  movel([0.337067, -0.804925, -2.801835, -1.105629, 1.570796, 1.907863],accel_mss,speed_ms,0,blend_radius_m)
  movel([0.336030, -0.804781, -2.801859, -1.105749, 1.570796, 1.906826],accel_mss,speed_ms,0,blend_radius_m)
  movel([0.330509, -0.802988, -2.802160, -1.107241, 1.570796, 1.901306],accel_mss,speed_ms,0,blend_radius_m)
  movel([0.325271, -0.800769, -2.802530, -1.109089, 1.570796, 1.896067],accel_mss,speed_ms,0,blend_radius_m)
  movel([0.320318, -0.798128, -2.802968, -1.111294, 1.570796, 1.891115],accel_mss,speed_ms,0,blend_radius_m)
  movel([0.315671, -0.795055, -2.803472, -1.113862, 1.570796, 1.886468],accel_mss,speed_ms,0,blend_radius_m)
  movel([0.314088, -0.793737, -2.803687, -1.114965, 1.570796, 1.884885],accel_mss,speed_ms,0,blend_radius_m)
  movel([0.312919, -0.791939, -2.803978, -1.116471, 1.570796, 1.883716],accel_mss,speed_ms,0,blend_radius_m)
  movel([0.312565, -0.790531, -2.804206, -1.117652, 1.570796, 1.883362],accel_mss,speed_ms,0,blend_radius_m)
  movel([0.312427, -0.788928, -2.804463, -1.118997, 1.570796, 1.883224],accel_mss,speed_ms,0,blend_radius_m)
  movel([0.312533, -0.785387, -2.805028, -1.121975, 1.570796, 1.883329],accel_mss,speed_ms,0,blend_radius_m)
  movel([0.314201, -0.771715, -2.807148, -1.133527, 1.570796, 1.884998],accel_mss,speed_ms,0,blend_radius_m)
  movel([0.314322, -0.768078, -2.807696, -1.136615, 1.570796, 1.885118],accel_mss,speed_ms,0,blend_radius_m)
  movel([0.313995, -0.765120, -2.808138, -1.139131, 1.570796, 1.884791],accel_mss,speed_ms,0,blend_radius_m)
  movel([0.313608, -0.764022, -2.808300, -1.140066, 1.570796, 1.884404],accel_mss,speed_ms,0,blend_radius_m)
  movel([0.313044, -0.763237, -2.808416, -1.140736, 1.570796, 1.883841],accel_mss,speed_ms,0,blend_radius_m)
  movel([0.312284, -0.762822, -2.808478, -1.141089, 1.570796, 1.883080],accel_mss,speed_ms,0,blend_radius_m)
  movel([0.311307, -0.762817, -2.808478, -1.141093, 1.570796, 1.882104],accel_mss,speed_ms,0,blend_radius_m)
  movel([0.309324, -0.763465, -2.808383, -1.140541, 1.570796, 1.880120],accel_mss,speed_ms,0,blend_radius_m)
  movel([0.308425, -0.763643, -2.808356, -1.140389, 1.570796, 1.879221],accel_mss,speed_ms,0,blend_radius_m)
  movel([0.307786, -0.763410, -2.808391, -1.140588, 1.570796, 1.878582],accel_mss,speed_ms,0,blend_radius_m)
  movel([0.307584, -0.762203, -2.808569, -1.141618, 1.570796, 1.878380],accel_mss,speed_ms,0,blend_radius_m)
  movel([0.307977, -0.760492, -2.808820, -1.143078, 1.570796, 1.878773],accel_mss,speed_ms,0,blend_radius_m)
  movel([0.309463, -0.754879, -2.809633, -1.147877, 1.570796, 1.880260],accel_mss,speed_ms,0,blend_radius_m)
  movel([0.310630, -0.749455, -2.810405, -1.152529, 1.570796, 1.881426],accel_mss,speed_ms,0,blend_radius_m)
  movel([0.312165, -0.739066, -2.811845, -1.161479, 1.570796, 1.882961],accel_mss,speed_ms,0,blend_radius_m)
  movel([0.312944, -0.729061, -2.813184, -1.170144, 1.570796, 1.883740],accel_mss,speed_ms,0,blend_radius_m)
  movel([0.313326, -0.719178, -2.814462, -1.178749, 1.570796, 1.884122],accel_mss,speed_ms,0,blend_radius_m)
  speed_ms = 0.005
  movel([0.313326, -0.711620, -2.807866, -1.192903, 1.570796, 1.884122],accel_mss,speed_ms,0,blend_radius_m)
  speed_ms = 0.040
  movel([0.305588, -0.730189, -2.805441, -1.176759, 1.570796, 1.876385],accel_mss,speed_ms,0,blend_radius_m)
  speed_ms = 0.005
  movel([0.305588, -0.737993, -2.811991, -1.162406, 1.570796, 1.876385],accel_mss,speed_ms,0,blend_radius_m)
  speed_ms = 0.025
  movel([0.301170, -0.750294, -2.810287, -1.151809, 1.570796, 1.871966],accel_mss,speed_ms,0,blend_radius_m)
  movel([0.298692, -0.756493, -2.809401, -1.146496, 1.570796, 1.869489],accel_mss,speed_ms,0,blend_radius_m)
  movel([0.296052, -0.762699, -2.808496, -1.141194, 1.570796, 1.866849],accel_mss,speed_ms,0,blend_radius_m)
  movel([0.293909, -0.761370, -2.808691, -1.142328, 1.570796, 1.864706],accel_mss,speed_ms,0,blend_radius_m)
  movel([0.293492, -0.761217, -2.808714, -1.142458, 1.570796, 1.864289],accel_mss,speed_ms,0,blend_radius_m)
  movel([0.292925, -0.761423, -2.808683, -1.142282, 1.570796, 1.863721],accel_mss,speed_ms,0,blend_radius_m)
  movel([0.292315, -0.762103, -2.808584, -1.141703, 1.570796, 1.863111],accel_mss,speed_ms,0,blend_radius_m)
  movel([0.291839, -0.762930, -2.808462, -1.140997, 1.570796, 1.862635],accel_mss,speed_ms,0,blend_radius_m)
  movel([0.288894, -0.768031, -2.807703, -1.136655, 1.570796, 1.859691],accel_mss,speed_ms,0,blend_radius_m)
  movel([0.285493, -0.772997, -2.806953, -1.132439, 1.570796, 1.856290],accel_mss,speed_ms,0,blend_radius_m)
  movel([0.284595, -0.774075, -2.806788, -1.131526, 1.570796, 1.855391],accel_mss,speed_ms,0,blend_radius_m)
  movel([0.283710, -0.774672, -2.806697, -1.131020, 1.570796, 1.854506],accel_mss,speed_ms,0,blend_radius_m)
  movel([0.283279, -0.774420, -2.806736, -1.131234, 1.570796, 1.854075],accel_mss,speed_ms,0,blend_radius_m)
  movel([0.283199, -0.773731, -2.806841, -1.131817, 1.570796, 1.853995],accel_mss,speed_ms,0,blend_radius_m)
  movel([0.283611, -0.768854, -2.807580, -1.135956, 1.570796, 1.854408],accel_mss,speed_ms,0,blend_radius_m)
  movel([0.284807, -0.763451, -2.808385, -1.140553, 1.570796, 1.855604],accel_mss,speed_ms,0,blend_radius_m)
  speed_ms = 0.005
  movel([0.284807, -0.755333, -2.801902, -1.155154, 1.570796, 1.855604],accel_mss,speed_ms,0,blend_radius_m)
  speed_ms = 0.040
  movel([0.290706, -0.762470, -2.800843, -1.149076, 1.570796, 1.861503],accel_mss,speed_ms,0,blend_radius_m)
  speed_ms = 0.005
  movel([0.290706, -0.770673, -2.807305, -1.134410, 1.570796, 1.861503],accel_mss,speed_ms,0,blend_radius_m)
  speed_ms = 0.025
  movel([0.289009, -0.778556, -2.806098, -1.127735, 1.570796, 1.859805],accel_mss,speed_ms,0,blend_radius_m)
  movel([0.287811, -0.782664, -2.805457, -1.124268, 1.570796, 1.858608],accel_mss,speed_ms,0,blend_radius_m)
  movel([0.284778, -0.791092, -2.804115, -1.117182, 1.570796, 1.855575],accel_mss,speed_ms,0,blend_radius_m)
  movel([0.282956, -0.795377, -2.803419, -1.113593, 1.570796, 1.853753],accel_mss,speed_ms,0,blend_radius_m)
  movel([0.278747, -0.803989, -2.801992, -1.106407, 1.570796, 1.849544],accel_mss,speed_ms,0,blend_radius_m)
  movel([0.279478, -0.801324, -2.802438, -1.108627, 1.570796, 1.850275],accel_mss,speed_ms,0,blend_radius_m)
  movel([0.279565, -0.799044, -2.802816, -1.110529, 1.570796, 1.850361],accel_mss,speed_ms,0,blend_radius_m)
  movel([0.279016, -0.797302, -2.803104, -1.111983, 1.570796, 1.849813],accel_mss,speed_ms,0,blend_radius_m)
  movel([0.277841, -0.796256, -2.803275, -1.112857, 1.570796, 1.848637],accel_mss,speed_ms,0,blend_radius_m)
  speed_ms = 0.005
  movel([0.277841, -0.787767, -2.796885, -1.127736, 1.570796, 1.848637],accel_mss,speed_ms,0,blend_radius_m)
  speed_ms = 0.040
  movel([0.251919, -0.805026, -2.793999, -1.113364, 1.570796, 1.822716],accel_mss,speed_ms,0,blend_radius_m)
  speed_ms = 0.005
  movel([0.251919, -0.813696, -2.800338, -1.098355, 1.570796, 1.822716],accel_mss,speed_ms,0,blend_radius_m)
  speed_ms = 0.025
  movel([0.247378, -0.819590, -2.799309, -1.093490, 1.570796, 1.818174],accel_mss,speed_ms,0,blend_radius_m)
  movel([0.242549, -0.825115, -2.798328, -1.088946, 1.570796, 1.813345],accel_mss,speed_ms,0,blend_radius_m)
  movel([0.237519, -0.830193, -2.797412, -1.084784, 1.570796, 1.808315],accel_mss,speed_ms,0,blend_radius_m)
  movel([0.232368, -0.834740, -2.796579, -1.081069, 1.570796, 1.803164],accel_mss,speed_ms,0,blend_radius_m)
  movel([0.233688, -0.832120, -2.797060, -1.083209, 1.570796, 1.804484],accel_mss,speed_ms,0,blend_radius_m)
  movel([0.234683, -0.829682, -2.797505, -1.085202, 1.570796, 1.805479],accel_mss,speed_ms,0,blend_radius_m)
  movel([0.235280, -0.827644, -2.797873, -1.086872, 1.570796, 1.806076],accel_mss,speed_ms,0,blend_radius_m)
  movel([0.235407, -0.826222, -2.798129, -1.088038, 1.570796, 1.806203],accel_mss,speed_ms,0,blend_radius_m)
  movel([0.234984, -0.825647, -2.798232, -1.088509, 1.570796, 1.805780],accel_mss,speed_ms,0,blend_radius_m)
  movel([0.234547, -0.825743, -2.798215, -1.088431, 1.570796, 1.805344],accel_mss,speed_ms,0,blend_radius_m)
  movel([0.233940, -0.826132, -2.798145, -1.088111, 1.570796, 1.804736],accel_mss,speed_ms,0,blend_radius_m)
  movel([0.232209, -0.827896, -2.797828, -1.086665, 1.570796, 1.803005],accel_mss,speed_ms,0,blend_radius_m)
  movel([0.227802, -0.833724, -2.796766, -1.081899, 1.570796, 1.798598],accel_mss,speed_ms,0,blend_radius_m)
  movel([0.225752, -0.836249, -2.796301, -1.079839, 1.570796, 1.796549],accel_mss,speed_ms,0,blend_radius_m)
  movel([0.221376, -0.840992, -2.795417, -1.075980, 1.570796, 1.792172],accel_mss,speed_ms,0,blend_radius_m)
  movel([0.219102, -0.843150, -2.795011, -1.074228, 1.570796, 1.789898],accel_mss,speed_ms,0,blend_radius_m)
  movel([0.216804, -0.845117, -2.794638, -1.072634, 1.570796, 1.787600],accel_mss,speed_ms,0,blend_radius_m)
  movel([0.214506, -0.846872, -2.794304, -1.071213, 1.570796, 1.785302],accel_mss,speed_ms,0,blend_radius_m)
  movel([0.212240, -0.848371, -2.794017, -1.070002, 1.570796, 1.783037],accel_mss,speed_ms,0,blend_radius_m)
  movel([0.215104, -0.844222, -2.794808, -1.073360, 1.570796, 1.785901],accel_mss,speed_ms,0,blend_radius_m)
  movel([0.217906, -0.840015, -2.795600, -1.076774, 1.570796, 1.788702],accel_mss,speed_ms,0,blend_radius_m)
  movel([0.219209, -0.837276, -2.796111, -1.079003, 1.570796, 1.790005],accel_mss,speed_ms,0,blend_radius_m)
  movel([0.219966, -0.834693, -2.796588, -1.081108, 1.570796, 1.790763],accel_mss,speed_ms,0,blend_radius_m)
  movel([0.219920, -0.833879, -2.796738, -1.081772, 1.570796, 1.790716],accel_mss,speed_ms,0,blend_radius_m)
  movel([0.219466, -0.833613, -2.796787, -1.081989, 1.570796, 1.790262],accel_mss,speed_ms,0,blend_radius_m)
  movel([0.218525, -0.834061, -2.796704, -1.081623, 1.570796, 1.789321],accel_mss,speed_ms,0,blend_radius_m)
  movel([0.217006, -0.835393, -2.796459, -1.080537, 1.570796, 1.787803],accel_mss,speed_ms,0,blend_radius_m)
  movel([0.209003, -0.843568, -2.794931, -1.073889, 1.570796, 1.779799],accel_mss,speed_ms,0,blend_radius_m)
  movel([0.205006, -0.847159, -2.794249, -1.070982, 1.570796, 1.775803],accel_mss,speed_ms,0,blend_radius_m)
  movel([0.203015, -0.848638, -2.793965, -1.069785, 1.570796, 1.773811],accel_mss,speed_ms,0,blend_radius_m)
  movel([0.201023, -0.849841, -2.793734, -1.068814, 1.570796, 1.771819],accel_mss,speed_ms,0,blend_radius_m)
  speed_ms = 0.005
  movel([0.201023, -0.840830, -2.787509, -1.084050, 1.570796, 1.771819],accel_mss,speed_ms,0,blend_radius_m)
  speed_ms = 0.040
  movel([0.238662, -0.785563, -2.797243, -1.129584, 1.570796, 1.809458],accel_mss,speed_ms,0,blend_radius_m)
  speed_ms = 0.005
  movel([0.238662, -0.794028, -2.803640, -1.114722, 1.570796, 1.809458],accel_mss,speed_ms,0,blend_radius_m)
  speed_ms = 0.025
  movel([0.238890, -0.790913, -2.804144, -1.117332, 1.570796, 1.809686],accel_mss,speed_ms,0,blend_radius_m)
  movel([0.239732, -0.787445, -2.804700, -1.120244, 1.570796, 1.810528],accel_mss,speed_ms,0,blend_radius_m)
  movel([0.241121, -0.783698, -2.805295, -1.123396, 1.570796, 1.811917],accel_mss,speed_ms,0,blend_radius_m)
  movel([0.242984, -0.779771, -2.805910, -1.126708, 1.570796, 1.813781],accel_mss,speed_ms,0,blend_radius_m)
  movel([0.245268, -0.775735, -2.806534, -1.130120, 1.570796, 1.816064],accel_mss,speed_ms,0,blend_radius_m)
  movel([0.247890, -0.771697, -2.807150, -1.133541, 1.570796, 1.818687],accel_mss,speed_ms,0,blend_radius_m)
  movel([0.250794, -0.767733, -2.807748, -1.136908, 1.570796, 1.821590],accel_mss,speed_ms,0,blend_radius_m)
  movel([0.253896, -0.763949, -2.808311, -1.140129, 1.570796, 1.824692],accel_mss,speed_ms,0,blend_radius_m)
  movel([0.257898, -0.759551, -2.808957, -1.143880, 1.570796, 1.828695],accel_mss,speed_ms,0,blend_radius_m)
  movel([0.266086, -0.750908, -2.810200, -1.151281, 1.570796, 1.836882],accel_mss,speed_ms,0,blend_radius_m)
  movel([0.270058, -0.746320, -2.810845, -1.155224, 1.570796, 1.840855],accel_mss,speed_ms,0,blend_radius_m)
  movel([0.273771, -0.741273, -2.811543, -1.159573, 1.570796, 1.844568],accel_mss,speed_ms,0,blend_radius_m)
  movel([0.275420, -0.738638, -2.811903, -1.161848, 1.570796, 1.846216],accel_mss,speed_ms,0,blend_radius_m)
  movel([0.276854, -0.736017, -2.812258, -1.164115, 1.570796, 1.847650],accel_mss,speed_ms,0,blend_radius_m)
  movel([0.278016, -0.733474, -2.812599, -1.166316, 1.570796, 1.848812],accel_mss,speed_ms,0,blend_radius_m)
  movel([0.278854, -0.731072, -2.812918, -1.168398, 1.570796, 1.849650],accel_mss,speed_ms,0,blend_radius_m)
  movel([0.279296, -0.728897, -2.813205, -1.170286, 1.570796, 1.850092],accel_mss,speed_ms,0,blend_radius_m)
  movel([0.279283, -0.727017, -2.813452, -1.171920, 1.570796, 1.850080],accel_mss,speed_ms,0,blend_radius_m)
  speed_ms = 0.005
  movel([0.279283, -0.719355, -2.806875, -1.186159, 1.570796, 1.850080],accel_mss,speed_ms,0,blend_radius_m)
  speed_ms = 0.040
  movel([0.278218, -0.705012, -2.808691, -1.198687, 1.570796, 1.849015],accel_mss,speed_ms,0,blend_radius_m)
  speed_ms = 0.005
  movel([0.278218, -0.712479, -2.815303, -1.184607, 1.570796, 1.849015],accel_mss,speed_ms,0,blend_radius_m)
  speed_ms = 0.025
  movel([0.274128, -0.726027, -2.813581, -1.172781, 1.570796, 1.844925],accel_mss,speed_ms,0,blend_radius_m)
  movel([0.272708, -0.729205, -2.813165, -1.170019, 1.570796, 1.843504],accel_mss,speed_ms,0,blend_radius_m)
  movel([0.270637, -0.732375, -2.812745, -1.167269, 1.570796, 1.841433],accel_mss,speed_ms,0,blend_radius_m)
  movel([0.268156, -0.735332, -2.812350, -1.164707, 1.570796, 1.838952],accel_mss,speed_ms,0,blend_radius_m)
  movel([0.259858, -0.744065, -2.811158, -1.157166, 1.570796, 1.830654],accel_mss,speed_ms,0,blend_radius_m)
  movel([0.257055, -0.747391, -2.810695, -1.154303, 1.570796, 1.827852],accel_mss,speed_ms,0,blend_radius_m)
  movel([0.254399, -0.750837, -2.810210, -1.151343, 1.570796, 1.825196],accel_mss,speed_ms,0,blend_radius_m)
  movel([0.251913, -0.754359, -2.809708, -1.148322, 1.570796, 1.822709],accel_mss,speed_ms,0,blend_radius_m)
  movel([0.249806, -0.757853, -2.809204, -1.145332, 1.570796, 1.820602],accel_mss,speed_ms,0,blend_radius_m)
  movel([0.248006, -0.761336, -2.808696, -1.142357, 1.570796, 1.818802],accel_mss,speed_ms,0,blend_radius_m)
  movel([0.246241, -0.764790, -2.808187, -1.139412, 1.570796, 1.817038],accel_mss,speed_ms,0,blend_radius_m)
  movel([0.244246, -0.768203, -2.807678, -1.136509, 1.570796, 1.815042],accel_mss,speed_ms,0,blend_radius_m)
  movel([0.242758, -0.762452, -2.808532, -1.141405, 1.570796, 1.813555],accel_mss,speed_ms,0,blend_radius_m)
  movel([0.243050, -0.760418, -2.808830, -1.143140, 1.570796, 1.813846],accel_mss,speed_ms,0,blend_radius_m)
  movel([0.243651, -0.758255, -2.809146, -1.144988, 1.570796, 1.814448],accel_mss,speed_ms,0,blend_radius_m)
  movel([0.244562, -0.755958, -2.809478, -1.146953, 1.570796, 1.815359],accel_mss,speed_ms,0,blend_radius_m)
  movel([0.245801, -0.753505, -2.809830, -1.149054, 1.570796, 1.816598],accel_mss,speed_ms,0,blend_radius_m)
  movel([0.248098, -0.750063, -2.810319, -1.152007, 1.570796, 1.818894],accel_mss,speed_ms,0,blend_radius_m)
  movel([0.251441, -0.745851, -2.810910, -1.155628, 1.570796, 1.822238],accel_mss,speed_ms,0,blend_radius_m)
  movel([0.259675, -0.736295, -2.812220, -1.163874, 1.570796, 1.830471],accel_mss,speed_ms,0,blend_radius_m)
  movel([0.263755, -0.731557, -2.812854, -1.167978, 1.570796, 1.834551],accel_mss,speed_ms,0,blend_radius_m)
  movel([0.267253, -0.727254, -2.813421, -1.171714, 1.570796, 1.838049],accel_mss,speed_ms,0,blend_radius_m)
  movel([0.269743, -0.723712, -2.813881, -1.174796, 1.570796, 1.840539],accel_mss,speed_ms,0,blend_radius_m)
  movel([0.270479, -0.722320, -2.814060, -1.176009, 1.570796, 1.841275],accel_mss,speed_ms,0,blend_radius_m)
  movel([0.270799, -0.721237, -2.814199, -1.176953, 1.570796, 1.841595],accel_mss,speed_ms,0,blend_radius_m)
  speed_ms = 0.005
  movel([0.270799, -0.713652, -2.807608, -1.191129, 1.570796, 1.841595],accel_mss,speed_ms,0,blend_radius_m)
  speed_ms = 0.040
  movel([0.256086, -0.716555, -2.807237, -1.188597, 1.570796, 1.826882],accel_mss,speed_ms,0,blend_radius_m)
  speed_ms = 0.005
  movel([0.256086, -0.724180, -2.813821, -1.174389, 1.570796, 1.826882],accel_mss,speed_ms,0,blend_radius_m)
  speed_ms = 0.025
  movel([0.254666, -0.724435, -2.813788, -1.174166, 1.570796, 1.825462],accel_mss,speed_ms,0,blend_radius_m)
  movel([0.253508, -0.724258, -2.813810, -1.174320, 1.570796, 1.824304],accel_mss,speed_ms,0,blend_radius_m)
  movel([0.251855, -0.722886, -2.813988, -1.175515, 1.570796, 1.822651],accel_mss,speed_ms,0,blend_radius_m)
  movel([0.250882, -0.720562, -2.814286, -1.177541, 1.570796, 1.821679],accel_mss,speed_ms,0,blend_radius_m)
  movel([0.250362, -0.717774, -2.814640, -1.179975, 1.570796, 1.821158],accel_mss,speed_ms,0,blend_radius_m)
  movel([0.250376, -0.716597, -2.814789, -1.181004, 1.570796, 1.821172],accel_mss,speed_ms,0,blend_radius_m)
  movel([0.251431, -0.714229, -2.815085, -1.183075, 1.570796, 1.822227],accel_mss,speed_ms,0,blend_radius_m)
  movel([0.255097, -0.707364, -2.815932, -1.189093, 1.570796, 1.825893],accel_mss,speed_ms,0,blend_radius_m)
  movel([0.261993, -0.693537, -2.817575, -1.201277, 1.570796, 1.832789],accel_mss,speed_ms,0,blend_radius_m)
  movel([0.265206, -0.686608, -2.818367, -1.207414, 1.570796, 1.836002],accel_mss,speed_ms,0,blend_radius_m)
  speed_ms = 0.005
  movel([0.265206, -0.679504, -2.811695, -1.221190, 1.570796, 1.836002],accel_mss,speed_ms,0,blend_radius_m)
  speed_ms = 0.040
  movel([0.255172, -0.687058, -2.810835, -1.214496, 1.570796, 1.825968],accel_mss,speed_ms,0,blend_radius_m)
  speed_ms = 0.005
  movel([0.255172, -0.694271, -2.817490, -1.200628, 1.570796, 1.825968],accel_mss,speed_ms,0,blend_radius_m)
  speed_ms = 0.025
  movel([0.253576, -0.698334, -2.817014, -1.197041, 1.570796, 1.824373],accel_mss,speed_ms,0,blend_radius_m)
  movel([0.251612, -0.702493, -2.816520, -1.193376, 1.570796, 1.822409],accel_mss,speed_ms,0,blend_radius_m)
  movel([0.249200, -0.706568, -2.816029, -1.189792, 1.570796, 1.819996],accel_mss,speed_ms,0,blend_radius_m)
  movel([0.247798, -0.708527, -2.815790, -1.188072, 1.570796, 1.818594],accel_mss,speed_ms,0,blend_radius_m)
  movel([0.244762, -0.712243, -2.815333, -1.184814, 1.570796, 1.815558],accel_mss,speed_ms,0,blend_radius_m)
  movel([0.243999, -0.713894, -2.815127, -1.183368, 1.570796, 1.814795],accel_mss,speed_ms,0,blend_radius_m)
  movel([0.239388, -0.726202, -2.813558, -1.172629, 1.570796, 1.810184],accel_mss,speed_ms,0,blend_radius_m)
  movel([0.238976, -0.727376, -2.813405, -1.171608, 1.570796, 1.809772],accel_mss,speed_ms,0,blend_radius_m)
  movel([0.238840, -0.728369, -2.813275, -1.170745, 1.570796, 1.809637],accel_mss,speed_ms,0,blend_radius_m)
  movel([0.239436, -0.729078, -2.813182, -1.170129, 1.570796, 1.810232],accel_mss,speed_ms,0,blend_radius_m)
  movel([0.240542, -0.729139, -2.813174, -1.170077, 1.570796, 1.811338],accel_mss,speed_ms,0,blend_radius_m)
  movel([0.243805, -0.729135, -2.813174, -1.170079, 1.570796, 1.814601],accel_mss,speed_ms,0,blend_radius_m)
  movel([0.246751, -0.729652, -2.813106, -1.169631, 1.570796, 1.817547],accel_mss,speed_ms,0,blend_radius_m)
  movel([0.249147, -0.730919, -2.812939, -1.168531, 1.570796, 1.819943],accel_mss,speed_ms,0,blend_radius_m)
  movel([0.250740, -0.733184, -2.812638, -1.166567, 1.570796, 1.821537],accel_mss,speed_ms,0,blend_radius_m)
  speed_ms = 0.005
  movel([0.250740, -0.725442, -2.806076, -1.180871, 1.570796, 1.821537],accel_mss,speed_ms,0,blend_radius_m)
  speed_ms = 0.040
  movel([0.239180, -0.756162, -2.801780, -1.154447, 1.570796, 1.809976],accel_mss,speed_ms,0,blend_radius_m)
  speed_ms = 0.005
  movel([0.239180, -0.764290, -2.808261, -1.139838, 1.570796, 1.809976],accel_mss,speed_ms,0,blend_radius_m)
  speed_ms = 0.025
  movel([0.238467, -0.765028, -2.808151, -1.139209, 1.570796, 1.809264],accel_mss,speed_ms,0,blend_radius_m)
  movel([0.237810, -0.765945, -2.808015, -1.138429, 1.570796, 1.808607],accel_mss,speed_ms,0,blend_radius_m)
  movel([0.235162, -0.770628, -2.807312, -1.134448, 1.570796, 1.805958],accel_mss,speed_ms,0,blend_radius_m)
  movel([0.234732, -0.771078, -2.807244, -1.134067, 1.570796, 1.805529],accel_mss,speed_ms,0,blend_radius_m)
  movel([0.234120, -0.771307, -2.807210, -1.133872, 1.570796, 1.804916],accel_mss,speed_ms,0,blend_radius_m)
  movel([0.233671, -0.771068, -2.807246, -1.134075, 1.570796, 1.804467],accel_mss,speed_ms,0,blend_radius_m)
  movel([0.233188, -0.769658, -2.807459, -1.135272, 1.570796, 1.803984],accel_mss,speed_ms,0,blend_radius_m)
  movel([0.233194, -0.766361, -2.807953, -1.138075, 1.570796, 1.803991],accel_mss,speed_ms,0,blend_radius_m)
  movel([0.234136, -0.762715, -2.808493, -1.141181, 1.570796, 1.804933],accel_mss,speed_ms,0,blend_radius_m)
  movel([0.235569, -0.758805, -2.809066, -1.144518, 1.570796, 1.806365],accel_mss,speed_ms,0,blend_radius_m)
  movel([0.237248, -0.754853, -2.809637, -1.147899, 1.570796, 1.808045],accel_mss,speed_ms,0,blend_radius_m)
  movel([0.239202, -0.750954, -2.810193, -1.151242, 1.570796, 1.809999],accel_mss,speed_ms,0,blend_radius_m)
  movel([0.241419, -0.747114, -2.810734, -1.154541, 1.570796, 1.812215],accel_mss,speed_ms,0,blend_radius_m)
  movel([0.243887, -0.743330, -2.811260, -1.157799, 1.570796, 1.814683],accel_mss,speed_ms,0,blend_radius_m)
  movel([0.246599, -0.739599, -2.811772, -1.161018, 1.570796, 1.817396],accel_mss,speed_ms,0,blend_radius_m)
  movel([0.249538, -0.735930, -2.812269, -1.164190, 1.570796, 1.820334],accel_mss,speed_ms,0,blend_radius_m)
  movel([0.252702, -0.732310, -2.812754, -1.167325, 1.570796, 1.823499],accel_mss,speed_ms,0,blend_radius_m)
  movel([0.256073, -0.728748, -2.813225, -1.170416, 1.570796, 1.826870],accel_mss,speed_ms,0,blend_radius_m)
  movel([0.260755, -0.723425, -2.813918, -1.175046, 1.570796, 1.831551],accel_mss,speed_ms,0,blend_radius_m)
  movel([0.265685, -0.717178, -2.814715, -1.180496, 1.570796, 1.836482],accel_mss,speed_ms,0,blend_radius_m)
  movel([0.271037, -0.709933, -2.815618, -1.186839, 1.570796, 1.841833],accel_mss,speed_ms,0,blend_radius_m)
  speed_ms = 0.005
  movel([0.271037, -0.702500, -2.808999, -1.200889, 1.570796, 1.841833],accel_mss,speed_ms,0,blend_radius_m)
  speed_ms = 0.040
  movel([0.266633, -0.704128, -2.808800, -1.199461, 1.570796, 1.837429],accel_mss,speed_ms,0,blend_radius_m)
  speed_ms = 0.005
  movel([0.266633, -0.711583, -2.815414, -1.185392, 1.570796, 1.837429],accel_mss,speed_ms,0,blend_radius_m)
  speed_ms = 0.025
  movel([0.271058, -0.701758, -2.816608, -1.194022, 1.570796, 1.841854],accel_mss,speed_ms,0,blend_radius_m)
  movel([0.275991, -0.691718, -2.817785, -1.202886, 1.570796, 1.846787],accel_mss,speed_ms,0,blend_radius_m)
  movel([0.278750, -0.686659, -2.818361, -1.207369, 1.570796, 1.849546],accel_mss,speed_ms,0,blend_radius_m)
  movel([0.281743, -0.681601, -2.818926, -1.211862, 1.570796, 1.852540],accel_mss,speed_ms,0,blend_radius_m)
  movel([0.285025, -0.676553, -2.819479, -1.216357, 1.570796, 1.855822],accel_mss,speed_ms,0,blend_radius_m)
  movel([0.288616, -0.671551, -2.820017, -1.220821, 1.570796, 1.859412],accel_mss,speed_ms,0,blend_radius_m)
  movel([0.298570, -0.659000, -2.821320, -1.232069, 1.570796, 1.869366],accel_mss,speed_ms,0,blend_radius_m)
  movel([0.302903, -0.653232, -2.821897, -1.237260, 1.570796, 1.873699],accel_mss,speed_ms,0,blend_radius_m)
  movel([0.304959, -0.650270, -2.822188, -1.239931, 1.570796, 1.875755],accel_mss,speed_ms,0,blend_radius_m)
  movel([0.306841, -0.647246, -2.822482, -1.242661, 1.570796, 1.877638],accel_mss,speed_ms,0,blend_radius_m)
  movel([0.311183, -0.638176, -2.823340, -1.250873, 1.570796, 1.881979],accel_mss,speed_ms,0,blend_radius_m)
  speed_ms = 0.005
  movel([0.311183, -0.631809, -2.816569, -1.264010, 1.570796, 1.881979],accel_mss,speed_ms,0,blend_radius_m)
  speed_ms = 0.040
  movel([0.321759, -0.610895, -2.818414, -1.283080, 1.570796, 1.892555],accel_mss,speed_ms,0,blend_radius_m)
  speed_ms = 0.005
  movel([0.321759, -0.616917, -2.825222, -1.270250, 1.570796, 1.892555],accel_mss,speed_ms,0,blend_radius_m)
  speed_ms = 0.025
  movel([0.325188, -0.609400, -2.825846, -1.277144, 1.570796, 1.895984],accel_mss,speed_ms,0,blend_radius_m)
  movel([0.327388, -0.605602, -2.826152, -1.280635, 1.570796, 1.898185],accel_mss,speed_ms,0,blend_radius_m)
  movel([0.330084, -0.601895, -2.826446, -1.284048, 1.570796, 1.900880],accel_mss,speed_ms,0,blend_radius_m)
  movel([0.332238, -0.599496, -2.826634, -1.286260, 1.570796, 1.903034],accel_mss,speed_ms,0,blend_radius_m)
  movel([0.334479, -0.597328, -2.826801, -1.288260, 1.570796, 1.905275],accel_mss,speed_ms,0,blend_radius_m)
  movel([0.339064, -0.593350, -2.827104, -1.291936, 1.570796, 1.909861],accel_mss,speed_ms,0,blend_radius_m)
  movel([0.343198, -0.589443, -2.827395, -1.295551, 1.570796, 1.913994],accel_mss,speed_ms,0,blend_radius_m)
  movel([0.346574, -0.585526, -2.827681, -1.299182, 1.570796, 1.917370],accel_mss,speed_ms,0,blend_radius_m)
  movel([0.353165, -0.576374, -2.828328, -1.307687, 1.570796, 1.923961],accel_mss,speed_ms,0,blend_radius_m)
  movel([0.354587, -0.574554, -2.828453, -1.309382, 1.570796, 1.925383],accel_mss,speed_ms,0,blend_radius_m)
  movel([0.356113, -0.572912, -2.828565, -1.310912, 1.570796, 1.926909],accel_mss,speed_ms,0,blend_radius_m)
  movel([0.359378, -0.570027, -2.828758, -1.313604, 1.570796, 1.930174],accel_mss,speed_ms,0,blend_radius_m)
  movel([0.365995, -0.564831, -2.829099, -1.318458, 1.570796, 1.936792],accel_mss,speed_ms,0,blend_radius_m)
  movel([0.373073, -0.558625, -2.829494, -1.324270, 1.570796, 1.943869],accel_mss,speed_ms,0,blend_radius_m)
  movel([0.376615, -0.555203, -2.829705, -1.327480, 1.570796, 1.947411],accel_mss,speed_ms,0,blend_radius_m)
  movel([0.380090, -0.551414, -2.829935, -1.331040, 1.570796, 1.950886],accel_mss,speed_ms,0,blend_radius_m)
  movel([0.382697, -0.548001, -2.830137, -1.334251, 1.570796, 1.953493],accel_mss,speed_ms,0,blend_radius_m)
  movel([0.384821, -0.544485, -2.830340, -1.337564, 1.570796, 1.955617],accel_mss,speed_ms,0,blend_radius_m)
  movel([0.385968, -0.541519, -2.830509, -1.340362, 1.570796, 1.956764],accel_mss,speed_ms,0,blend_radius_m)
  movel([0.386018, -0.540452, -2.830568, -1.341368, 1.570796, 1.956814],accel_mss,speed_ms,0,blend_radius_m)
  movel([0.385633, -0.539775, -2.830606, -1.342008, 1.570796, 1.956430],accel_mss,speed_ms,0,blend_radius_m)
  movel([0.384024, -0.539347, -2.830630, -1.342412, 1.570796, 1.954820],accel_mss,speed_ms,0,blend_radius_m)
  movel([0.381703, -0.539729, -2.830609, -1.342051, 1.570796, 1.952500],accel_mss,speed_ms,0,blend_radius_m)
  movel([0.378837, -0.540820, -2.830548, -1.341021, 1.570796, 1.949633],accel_mss,speed_ms,0,blend_radius_m)
  movel([0.375629, -0.542477, -2.830455, -1.339457, 1.570796, 1.946425],accel_mss,speed_ms,0,blend_radius_m)
  movel([0.372254, -0.544602, -2.830334, -1.337453, 1.570796, 1.943051],accel_mss,speed_ms,0,blend_radius_m)
  movel([0.368906, -0.547056, -2.830192, -1.335142, 1.570796, 1.939702],accel_mss,speed_ms,0,blend_radius_m)
  movel([0.365765, -0.549727, -2.830035, -1.332627, 1.570796, 1.936562],accel_mss,speed_ms,0,blend_radius_m)
  movel([0.363011, -0.552495, -2.829870, -1.330024, 1.570796, 1.933807],accel_mss,speed_ms,0,blend_radius_m)
  movel([0.359228, -0.557153, -2.829585, -1.325651, 1.570796, 1.930024],accel_mss,speed_ms,0,blend_radius_m)
  movel([0.348676, -0.571461, -2.828662, -1.312265, 1.570796, 1.919472],accel_mss,speed_ms,0,blend_radius_m)
  movel([0.341420, -0.580615, -2.828032, -1.303742, 1.570796, 1.912216],accel_mss,speed_ms,0,blend_radius_m)
  movel([0.334837, -0.587979, -2.827503, -1.296907, 1.570796, 1.905633],accel_mss,speed_ms,0,blend_radius_m)
  movel([0.331585, -0.591547, -2.827239, -1.293603, 1.570796, 1.902381],accel_mss,speed_ms,0,blend_radius_m)
  movel([0.328499, -0.595253, -2.826960, -1.290176, 1.570796, 1.899296],accel_mss,speed_ms,0,blend_radius_m)
  movel([0.325566, -0.599275, -2.826651, -1.286464, 1.570796, 1.896362],accel_mss,speed_ms,0,blend_radius_m)
  movel([0.322921, -0.603318, -2.826334, -1.282737, 1.570796, 1.893717],accel_mss,speed_ms,0,blend_radius_m)
  movel([0.320533, -0.607368, -2.826010, -1.279011, 1.570796, 1.891330],accel_mss,speed_ms,0,blend_radius_m)
  movel([0.318373, -0.611394, -2.825682, -1.275313, 1.570796, 1.889170],accel_mss,speed_ms,0,blend_radius_m)
  movel([0.314600, -0.619311, -2.825019, -1.268059, 1.570796, 1.885397],accel_mss,speed_ms,0,blend_radius_m)
  movel([0.311326, -0.626923, -2.824358, -1.261108, 1.570796, 1.882122],accel_mss,speed_ms,0,blend_radius_m)
  speed_ms = 0.005
  movel([0.311326, -0.620737, -2.817568, -1.274084, 1.570796, 1.882122],accel_mss,speed_ms,0,blend_radius_m)
  speed_ms = 0.040
  movel([0.303174, -0.627998, -2.816919, -1.267472, 1.570796, 1.873970],accel_mss,speed_ms,0,blend_radius_m)
  speed_ms = 0.005
  movel([0.303174, -0.634303, -2.823696, -1.254390, 1.570796, 1.873970],accel_mss,speed_ms,0,blend_radius_m)
  speed_ms = 0.025
  movel([0.308567, -0.622268, -2.824765, -1.265356, 1.570796, 1.879363],accel_mss,speed_ms,0,blend_radius_m)
  movel([0.311017, -0.617155, -2.825202, -1.270032, 1.570796, 1.881813],accel_mss,speed_ms,0,blend_radius_m)
  movel([0.313262, -0.612099, -2.825624, -1.274666, 1.570796, 1.884058],accel_mss,speed_ms,0,blend_radius_m)
  movel([0.314771, -0.607909, -2.825967, -1.278513, 1.570796, 1.885567],accel_mss,speed_ms,0,blend_radius_m)
  movel([0.315798, -0.603986, -2.826281, -1.282122, 1.570796, 1.886594],accel_mss,speed_ms,0,blend_radius_m)
  movel([0.316319, -0.600410, -2.826562, -1.285417, 1.570796, 1.887116],accel_mss,speed_ms,0,blend_radius_m)
  movel([0.316316, -0.597266, -2.826806, -1.288318, 1.570796, 1.887112],accel_mss,speed_ms,0,blend_radius_m)
  movel([0.318007, -0.595920, -2.826909, -1.289560, 1.570796, 1.888803],accel_mss,speed_ms,0,blend_radius_m)
  movel([0.319623, -0.594979, -2.826980, -1.290430, 1.570796, 1.890419],accel_mss,speed_ms,0,blend_radius_m)
  movel([0.322733, -0.593608, -2.827084, -1.291696, 1.570796, 1.893529],accel_mss,speed_ms,0,blend_radius_m)
  movel([0.326035, -0.591866, -2.827215, -1.293308, 1.570796, 1.896831],accel_mss,speed_ms,0,blend_radius_m)
  movel([0.327738, -0.590557, -2.827313, -1.294519, 1.570796, 1.898535],accel_mss,speed_ms,0,blend_radius_m)
  movel([0.329386, -0.588811, -2.827442, -1.296137, 1.570796, 1.900182],accel_mss,speed_ms,0,blend_radius_m)
  movel([0.348272, -0.565665, -2.829045, -1.317679, 1.570796, 1.919069],accel_mss,speed_ms,0,blend_radius_m)
  movel([0.348583, -0.563195, -2.829205, -1.319989, 1.570796, 1.919380],accel_mss,speed_ms,0,blend_radius_m)
  movel([0.348124, -0.561343, -2.829323, -1.321723, 1.570796, 1.918921],accel_mss,speed_ms,0,blend_radius_m)
  movel([0.346919, -0.560208, -2.829395, -1.322787, 1.570796, 1.917716],accel_mss,speed_ms,0,blend_radius_m)
  movel([0.345019, -0.559872, -2.829416, -1.323101, 1.570796, 1.915815],accel_mss,speed_ms,0,blend_radius_m)
  movel([0.348929, -0.557437, -2.829568, -1.325384, 1.570796, 1.919726],accel_mss,speed_ms,0,blend_radius_m)
  movel([0.352511, -0.555837, -2.829667, -1.326885, 1.570796, 1.923308],accel_mss,speed_ms,0,blend_radius_m)
  movel([0.355579, -0.555141, -2.829709, -1.327539, 1.570796, 1.926375],accel_mss,speed_ms,0,blend_radius_m)
  movel([0.357960, -0.555407, -2.829693, -1.327289, 1.570796, 1.928756],accel_mss,speed_ms,0,blend_radius_m)
  speed_ms = 0.005
  movel([0.357960, -0.550452, -2.822792, -1.339144, 1.570796, 1.928756],accel_mss,speed_ms,0,blend_radius_m)
  speed_ms = 0.040
  movel([0.361776, -0.539696, -2.823428, -1.349265, 1.570796, 1.932572],accel_mss,speed_ms,0,blend_radius_m)
  speed_ms = 0.005
  movel([0.361776, -0.544451, -2.830342, -1.337596, 1.570796, 1.932572],accel_mss,speed_ms,0,blend_radius_m)
  speed_ms = 0.025
  movel([0.364576, -0.538316, -2.830687, -1.343386, 1.570796, 1.935373],accel_mss,speed_ms,0,blend_radius_m)
  movel([0.366892, -0.532590, -2.830996, -1.348802, 1.570796, 1.937688],accel_mss,speed_ms,0,blend_radius_m)
  movel([0.368755, -0.527230, -2.831276, -1.353883, 1.570796, 1.939551],accel_mss,speed_ms,0,blend_radius_m)
  movel([0.370195, -0.522193, -2.831529, -1.358667, 1.570796, 1.940991],accel_mss,speed_ms,0,blend_radius_m)
  movel([0.371243, -0.517429, -2.831760, -1.363200, 1.570796, 1.942039],accel_mss,speed_ms,0,blend_radius_m)
  movel([0.371933, -0.512886, -2.831973, -1.367530, 1.570796, 1.942730],accel_mss,speed_ms,0,blend_radius_m)
  movel([0.372379, -0.504267, -2.832357, -1.375764, 1.570796, 1.943176],accel_mss,speed_ms,0,blend_radius_m)
  movel([0.362866, -0.525432, -2.831367, -1.355590, 1.570796, 1.933663],accel_mss,speed_ms,0,blend_radius_m)
  movel([0.363724, -0.523187, -2.831480, -1.357723, 1.570796, 1.934521],accel_mss,speed_ms,0,blend_radius_m)
  movel([0.364223, -0.521167, -2.831579, -1.359643, 1.570796, 1.935019],accel_mss,speed_ms,0,blend_radius_m)
  movel([0.364264, -0.517768, -2.831744, -1.362877, 1.570796, 1.935060],accel_mss,speed_ms,0,blend_radius_m)
  movel([0.363219, -0.515170, -2.831867, -1.365352, 1.570796, 1.934016],accel_mss,speed_ms,0,blend_radius_m)
  movel([0.361350, -0.513295, -2.831954, -1.367140, 1.570796, 1.932147],accel_mss,speed_ms,0,blend_radius_m)
  movel([0.358908, -0.512054, -2.832011, -1.368324, 1.570796, 1.929705],accel_mss,speed_ms,0,blend_radius_m)
  movel([0.356160, -0.511362, -2.832043, -1.368984, 1.570796, 1.926956],accel_mss,speed_ms,0,blend_radius_m)
  movel([0.350805, -0.511242, -2.832048, -1.369099, 1.570796, 1.921601],accel_mss,speed_ms,0,blend_radius_m)
  movel([0.352322, -0.517338, -2.831764, -1.363287, 1.570796, 1.923118],accel_mss,speed_ms,0,blend_radius_m)
  movel([0.352350, -0.521152, -2.831580, -1.359657, 1.570796, 1.923146],accel_mss,speed_ms,0,blend_radius_m)
  movel([0.351411, -0.525467, -2.831365, -1.355557, 1.570796, 1.922207],accel_mss,speed_ms,0,blend_radius_m)
  movel([0.349024, -0.526346, -2.831321, -1.354722, 1.570796, 1.919820],accel_mss,speed_ms,0,blend_radius_m)
  movel([0.346872, -0.526693, -2.831303, -1.354393, 1.570796, 1.917668],accel_mss,speed_ms,0,blend_radius_m)
  movel([0.342914, -0.526512, -2.831312, -1.354565, 1.570796, 1.913711],accel_mss,speed_ms,0,blend_radius_m)
  movel([0.338862, -0.526325, -2.831322, -1.354742, 1.570796, 1.909658],accel_mss,speed_ms,0,blend_radius_m)
  movel([0.336592, -0.526665, -2.831305, -1.354419, 1.570796, 1.907388],accel_mss,speed_ms,0,blend_radius_m)
  movel([0.334061, -0.527515, -2.831261, -1.353613, 1.570796, 1.904857],accel_mss,speed_ms,0,blend_radius_m)
  movel([0.331141, -0.533123, -2.830968, -1.348298, 1.570796, 1.901938],accel_mss,speed_ms,0,blend_radius_m)
  movel([0.329142, -0.538316, -2.830687, -1.343386, 1.570796, 1.899939],accel_mss,speed_ms,0,blend_radius_m)
  movel([0.325579, -0.539995, -2.830594, -1.341800, 1.570796, 1.896375],accel_mss,speed_ms,0,blend_radius_m)
  movel([0.322366, -0.540955, -2.830540, -1.340894, 1.570796, 1.893163],accel_mss,speed_ms,0,blend_radius_m)
  movel([0.319565, -0.541176, -2.830528, -1.340685, 1.570796, 1.890361],accel_mss,speed_ms,0,blend_radius_m)
  movel([0.317254, -0.540651, -2.830557, -1.341181, 1.570796, 1.888051],accel_mss,speed_ms,0,blend_radius_m)
  movel([0.316801, -0.541261, -2.830523, -1.340605, 1.570796, 1.887598],accel_mss,speed_ms,0,blend_radius_m)
  movel([0.312948, -0.548274, -2.830121, -1.333995, 1.570796, 1.883744],accel_mss,speed_ms,0,blend_radius_m)
  movel([0.308518, -0.556883, -2.829602, -1.325904, 1.570796, 1.879314],accel_mss,speed_ms,0,blend_radius_m)
  movel([0.306832, -0.560869, -2.829353, -1.322167, 1.570796, 1.877628],accel_mss,speed_ms,0,blend_radius_m)
  movel([0.305575, -0.564420, -2.829126, -1.318843, 1.570796, 1.876371],accel_mss,speed_ms,0,blend_radius_m)
  movel([0.303731, -0.571374, -2.828668, -1.312346, 1.570796, 1.874527],accel_mss,speed_ms,0,blend_radius_m)
  movel([0.296179, -0.567959, -2.828895, -1.315535, 1.570796, 1.866975],accel_mss,speed_ms,0,blend_radius_m)
  movel([0.294293, -0.572174, -2.828614, -1.311600, 1.570796, 1.865090],accel_mss,speed_ms,0,blend_radius_m)
  movel([0.292708, -0.576277, -2.828335, -1.307777, 1.570796, 1.863505],accel_mss,speed_ms,0,blend_radius_m)
  movel([0.290333, -0.584107, -2.827784, -1.300498, 1.570796, 1.861129],accel_mss,speed_ms,0,blend_radius_m)
  movel([0.288921, -0.591285, -2.827258, -1.293846, 1.570796, 1.859717],accel_mss,speed_ms,0,blend_radius_m)
  movel([0.288123, -0.599624, -2.826624, -1.286141, 1.570796, 1.858919],accel_mss,speed_ms,0,blend_radius_m)
  movel([0.287779, -0.600740, -2.826537, -1.285113, 1.570796, 1.858575],accel_mss,speed_ms,0,blend_radius_m)
  movel([0.287159, -0.601956, -2.826441, -1.283992, 1.570796, 1.857956],accel_mss,speed_ms,0,blend_radius_m)
  movel([0.285929, -0.603566, -2.826314, -1.282509, 1.570796, 1.856725],accel_mss,speed_ms,0,blend_radius_m)
  movel([0.276804, -0.612653, -2.825578, -1.274158, 1.570796, 1.847600],accel_mss,speed_ms,0,blend_radius_m)
  movel([0.272177, -0.616657, -2.825244, -1.270488, 1.570796, 1.842973],accel_mss,speed_ms,0,blend_radius_m)
  movel([0.270488, -0.617741, -2.825153, -1.269496, 1.570796, 1.841284],accel_mss,speed_ms,0,blend_radius_m)
  movel([0.269521, -0.617847, -2.825144, -1.269399, 1.570796, 1.840317],accel_mss,speed_ms,0,blend_radius_m)
  movel([0.273197, -0.620149, -2.824947, -1.267293, 1.570796, 1.843994],accel_mss,speed_ms,0,blend_radius_m)
  movel([0.275377, -0.620824, -2.824890, -1.266675, 1.570796, 1.846174],accel_mss,speed_ms,0,blend_radius_m)
  movel([0.277763, -0.621187, -2.824858, -1.266343, 1.570796, 1.848560],accel_mss,speed_ms,0,blend_radius_m)
  movel([0.269994, -0.631437, -2.823956, -1.256997, 1.570796, 1.840790],accel_mss,speed_ms,0,blend_radius_m)
  movel([0.261856, -0.642689, -2.822917, -1.246783, 1.570796, 1.832652],accel_mss,speed_ms,0,blend_radius_m)
  movel([0.258032, -0.648356, -2.822374, -1.241658, 1.570796, 1.828829],accel_mss,speed_ms,0,blend_radius_m)
  movel([0.254566, -0.653869, -2.821834, -1.236686, 1.570796, 1.825362],accel_mss,speed_ms,0,blend_radius_m)
  movel([0.251604, -0.659107, -2.821309, -1.231973, 1.570796, 1.822400],accel_mss,speed_ms,0,blend_radius_m)
  movel([0.249284, -0.663940, -2.820815, -1.227634, 1.570796, 1.820080],accel_mss,speed_ms,0,blend_radius_m)
  movel([0.252859, -0.660132, -2.821205, -1.231052, 1.570796, 1.823656],accel_mss,speed_ms,0,blend_radius_m)
  movel([0.256515, -0.656621, -2.821560, -1.234208, 1.570796, 1.827311],accel_mss,speed_ms,0,blend_radius_m)
  movel([0.260205, -0.653484, -2.821872, -1.237033, 1.570796, 1.831001],accel_mss,speed_ms,0,blend_radius_m)
  movel([0.263905, -0.650786, -2.822138, -1.239465, 1.570796, 1.834702],accel_mss,speed_ms,0,blend_radius_m)
  movel([0.261399, -0.653851, -2.821836, -1.236702, 1.570796, 1.832196],accel_mss,speed_ms,0,blend_radius_m)
  movel([0.256818, -0.660213, -2.821197, -1.230979, 1.570796, 1.827614],accel_mss,speed_ms,0,blend_radius_m)
  movel([0.254774, -0.663458, -2.820865, -1.228067, 1.570796, 1.825570],accel_mss,speed_ms,0,blend_radius_m)
  movel([0.251273, -0.669892, -2.820193, -1.222304, 1.570796, 1.822070],accel_mss,speed_ms,0,blend_radius_m)
  movel([0.249845, -0.673034, -2.819859, -1.219496, 1.570796, 1.820641],accel_mss,speed_ms,0,blend_radius_m)
  movel([0.248659, -0.676078, -2.819531, -1.216780, 1.570796, 1.819455],accel_mss,speed_ms,0,blend_radius_m)
  speed_ms = 0.005
  movel([0.248659, -0.669128, -2.812837, -1.230424, 1.570796, 1.819455],accel_mss,speed_ms,0,blend_radius_m)
  speed_ms = 0.040
  movel([0.261096, -0.670341, -2.812706, -1.229343, 1.570796, 1.831893],accel_mss,speed_ms,0,blend_radius_m)
  speed_ms = 0.005
  movel([0.261096, -0.677309, -2.819397, -1.215683, 1.570796, 1.831893],accel_mss,speed_ms,0,blend_radius_m)
  speed_ms = 0.025
  movel([0.261978, -0.673487, -2.819810, -1.219092, 1.570796, 1.832775],accel_mss,speed_ms,0,blend_radius_m)
  movel([0.263180, -0.669438, -2.820241, -1.222710, 1.570796, 1.833976],accel_mss,speed_ms,0,blend_radius_m)
  movel([0.264694, -0.665200, -2.820685, -1.226505, 1.570796, 1.835491],accel_mss,speed_ms,0,blend_radius_m)
  movel([0.266514, -0.660816, -2.821136, -1.230437, 1.570796, 1.837310],accel_mss,speed_ms,0,blend_radius_m)
  movel([0.268640, -0.656317, -2.821590, -1.234482, 1.570796, 1.839436],accel_mss,speed_ms,0,blend_radius_m)
  movel([0.271058, -0.651746, -2.822044, -1.238600, 1.570796, 1.841854],accel_mss,speed_ms,0,blend_radius_m)
  movel([0.273763, -0.647137, -2.822492, -1.242759, 1.570796, 1.844560],accel_mss,speed_ms,0,blend_radius_m)
  movel([0.276750, -0.642538, -2.822931, -1.246920, 1.570796, 1.847547],accel_mss,speed_ms,0,blend_radius_m)
  movel([0.286612, -0.628210, -2.824244, -1.259935, 1.570796, 1.857408],accel_mss,speed_ms,0,blend_radius_m)
  movel([0.288661, -0.624853, -2.824540, -1.262995, 1.570796, 1.859457],accel_mss,speed_ms,0,blend_radius_m)
  movel([0.290516, -0.621419, -2.824838, -1.266132, 1.570796, 1.861312],accel_mss,speed_ms,0,blend_radius_m)
  movel([0.292163, -0.617829, -2.825145, -1.269415, 1.570796, 1.862959],accel_mss,speed_ms,0,blend_radius_m)
  movel([0.293595, -0.613989, -2.825468, -1.272932, 1.570796, 1.864391],accel_mss,speed_ms,0,blend_radius_m)
  movel([0.296721, -0.603369, -2.826330, -1.282690, 1.570796, 1.867517],accel_mss,speed_ms,0,blend_radius_m)
  movel([0.298529, -0.597930, -2.826755, -1.287704, 1.570796, 1.869326],accel_mss,speed_ms,0,blend_radius_m)
  movel([0.301036, -0.592150, -2.827194, -1.293045, 1.570796, 1.871832],accel_mss,speed_ms,0,blend_radius_m)
  movel([0.303004, -0.588498, -2.827465, -1.296426, 1.570796, 1.873800],accel_mss,speed_ms,0,blend_radius_m)
  movel([0.305252, -0.584823, -2.827732, -1.299834, 1.570796, 1.876048],accel_mss,speed_ms,0,blend_radius_m)
  movel([0.310421, -0.577459, -2.828253, -1.306677, 1.570796, 1.881218],accel_mss,speed_ms,0,blend_radius_m)
  movel([0.316191, -0.570138, -2.828751, -1.313500, 1.570796, 1.886988],accel_mss,speed_ms,0,blend_radius_m)
  movel([0.322221, -0.562941, -2.829221, -1.320226, 1.570796, 1.893018],accel_mss,speed_ms,0,blend_radius_m)
  movel([0.328174, -0.556066, -2.829652, -1.326671, 1.570796, 1.898970],accel_mss,speed_ms,0,blend_radius_m)
  movel([0.334338, -0.549476, -2.830050, -1.332864, 1.570796, 1.905134],accel_mss,speed_ms,0,blend_radius_m)
  movel([0.337426, -0.546499, -2.830224, -1.335665, 1.570796, 1.908222],accel_mss,speed_ms,0,blend_radius_m)
  movel([0.340487, -0.543837, -2.830377, -1.338175, 1.570796, 1.911284],accel_mss,speed_ms,0,blend_radius_m)
  movel([0.343472, -0.541594, -2.830504, -1.340291, 1.570796, 1.914269],accel_mss,speed_ms,0,blend_radius_m)
  movel([0.346372, -0.539832, -2.830603, -1.341954, 1.570796, 1.917168],accel_mss,speed_ms,0,blend_radius_m)
  speed_ms = 0.005
  movel([0.346372, -0.535163, -2.823683, -1.353543, 1.570796, 1.917168],accel_mss,speed_ms,0,blend_radius_m)
  speed_ms = 0.040
  movel([0.349211, -0.536682, -2.823599, -1.352108, 1.570796, 1.920007],accel_mss,speed_ms,0,blend_radius_m)
  speed_ms = 0.005
  movel([0.349211, -0.541381, -2.830516, -1.340492, 1.570796, 1.920007],accel_mss,speed_ms,0,blend_radius_m)
  speed_ms = 0.025
  movel([0.350136, -0.541721, -2.830497, -1.340171, 1.570796, 1.920932],accel_mss,speed_ms,0,blend_radius_m)
  movel([0.351314, -0.542509, -2.830453, -1.339428, 1.570796, 1.922110],accel_mss,speed_ms,0,blend_radius_m)
  movel([0.352745, -0.545735, -2.830268, -1.336385, 1.570796, 1.923541],accel_mss,speed_ms,0,blend_radius_m)
  movel([0.352995, -0.547851, -2.830145, -1.334393, 1.570796, 1.923791],accel_mss,speed_ms,0,blend_radius_m)
  movel([0.352756, -0.549134, -2.830070, -1.333185, 1.570796, 1.923552],accel_mss,speed_ms,0,blend_radius_m)
  movel([0.352424, -0.549546, -2.830046, -1.332797, 1.570796, 1.923220],accel_mss,speed_ms,0,blend_radius_m)
  movel([0.351896, -0.549703, -2.830036, -1.332649, 1.570796, 1.922692],accel_mss,speed_ms,0,blend_radius_m)
  movel([0.346949, -0.549394, -2.830055, -1.332940, 1.570796, 1.917745],accel_mss,speed_ms,0,blend_radius_m)
  movel([0.344047, -0.549947, -2.830022, -1.332420, 1.570796, 1.914843],accel_mss,speed_ms,0,blend_radius_m)
  movel([0.342393, -0.550684, -2.829978, -1.331727, 1.570796, 1.913189],accel_mss,speed_ms,0,blend_radius_m)
  movel([0.340568, -0.551820, -2.829910, -1.330659, 1.570796, 1.911364],accel_mss,speed_ms,0,blend_radius_m)
  movel([0.338416, -0.553571, -2.829805, -1.329013, 1.570796, 1.909212],accel_mss,speed_ms,0,blend_radius_m)
  movel([0.336248, -0.555618, -2.829680, -1.327091, 1.570796, 1.907045],accel_mss,speed_ms,0,blend_radius_m)
  movel([0.330981, -0.561061, -2.829341, -1.321988, 1.570796, 1.901778],accel_mss,speed_ms,0,blend_radius_m)
  movel([0.325797, -0.566917, -2.828964, -1.316509, 1.570796, 1.896593],accel_mss,speed_ms,0,blend_radius_m)
  movel([0.320854, -0.572999, -2.828559, -1.310831, 1.570796, 1.891650],accel_mss,speed_ms,0,blend_radius_m)
  movel([0.316321, -0.579099, -2.828139, -1.305151, 1.570796, 1.887118],accel_mss,speed_ms,0,blend_radius_m)
  movel([0.318210, -0.583504, -2.827827, -1.301058, 1.570796, 1.889007],accel_mss,speed_ms,0,blend_radius_m)
  movel([0.319268, -0.588764, -2.827445, -1.296180, 1.570796, 1.890065],accel_mss,speed_ms,0,blend_radius_m)
  movel([0.317463, -0.588522, -2.827463, -1.296404, 1.570796, 1.888260],accel_mss,speed_ms,0,blend_radius_m)
  movel([0.315279, -0.588916, -2.827434, -1.296039, 1.570796, 1.886076],accel_mss,speed_ms,0,blend_radius_m)
  movel([0.312783, -0.589941, -2.827358, -1.295090, 1.570796, 1.883579],accel_mss,speed_ms,0,blend_radius_m)
  movel([0.310067, -0.591555, -2.827238, -1.293596, 1.570796, 1.880864],accel_mss,speed_ms,0,blend_radius_m)
  movel([0.308732, -0.592765, -2.827148, -1.292477, 1.570796, 1.879528],accel_mss,speed_ms,0,blend_radius_m)
  movel([0.308074, -0.594133, -2.827045, -1.291211, 1.570796, 1.878870],accel_mss,speed_ms,0,blend_radius_m)
  movel([0.303568, -0.607872, -2.825970, -1.278547, 1.570796, 1.874364],accel_mss,speed_ms,0,blend_radius_m)
  movel([0.300842, -0.615035, -2.825380, -1.271974, 1.570796, 1.871639],accel_mss,speed_ms,0,blend_radius_m)
  movel([0.297673, -0.622460, -2.824749, -1.265181, 1.570796, 1.868470],accel_mss,speed_ms,0,blend_radius_m)
  movel([0.294091, -0.629963, -2.824088, -1.258338, 1.570796, 1.864887],accel_mss,speed_ms,0,blend_radius_m)
  movel([0.290108, -0.637383, -2.823413, -1.251593, 1.570796, 1.860904],accel_mss,speed_ms,0,blend_radius_m)
  movel([0.281824, -0.652228, -2.821996, -1.238165, 1.570796, 1.852621],accel_mss,speed_ms,0,blend_radius_m)
  movel([0.278355, -0.659377, -2.821282, -1.231730, 1.570796, 1.849151],accel_mss,speed_ms,0,blend_radius_m)
  movel([0.275692, -0.666307, -2.820569, -1.225512, 1.570796, 1.846488],accel_mss,speed_ms,0,blend_radius_m)
  speed_ms = 0.005
  movel([0.275692, -0.659504, -2.813855, -1.239031, 1.570796, 1.846488],accel_mss,speed_ms,0,blend_radius_m)
  speed_ms = 0.040
  movel([0.303078, -0.639490, -2.815848, -1.257051, 1.570796, 1.873874],accel_mss,speed_ms,0,blend_radius_m)
  speed_ms = 0.005
  movel([0.303078, -0.645980, -2.822603, -1.243805, 1.570796, 1.873874],accel_mss,speed_ms,0,blend_radius_m)
  speed_ms = 0.025
  movel([0.300877, -0.651656, -2.822052, -1.238681, 1.570796, 1.871673],accel_mss,speed_ms,0,blend_radius_m)
  movel([0.297944, -0.657558, -2.821466, -1.233366, 1.570796, 1.868740],accel_mss,speed_ms,0,blend_radius_m)
  movel([0.294388, -0.663483, -2.820862, -1.228044, 1.570796, 1.865184],accel_mss,speed_ms,0,blend_radius_m)
  movel([0.290325, -0.669245, -2.820261, -1.222882, 1.570796, 1.861122],accel_mss,speed_ms,0,blend_radius_m)
  speed_ms = 0.005
  movel([0.290325, -0.662397, -2.813553, -1.236439, 1.570796, 1.861122],accel_mss,speed_ms,0,blend_radius_m)
  speed_ms = 0.040
  movel([0.285559, -0.658387, -2.813970, -1.240032, 1.570796, 1.856356],accel_mss,speed_ms,0,blend_radius_m)
  speed_ms = 0.005
  movel([0.285559, -0.665173, -2.820687, -1.226528, 1.570796, 1.856356],accel_mss,speed_ms,0,blend_radius_m)
  speed_ms = 0.025
  movel([0.265122, -0.701697, -2.816615, -1.194076, 1.570796, 1.835919],accel_mss,speed_ms,0,blend_radius_m)
  movel([0.264110, -0.703940, -2.816347, -1.192103, 1.570796, 1.834906],accel_mss,speed_ms,0,blend_radius_m)
  movel([0.264152, -0.705969, -2.816102, -1.190318, 1.570796, 1.834948],accel_mss,speed_ms,0,blend_radius_m)
  movel([0.264198, -0.708590, -2.815782, -1.188016, 1.570796, 1.834995],accel_mss,speed_ms,0,blend_radius_m)
  movel([0.263580, -0.711699, -2.815400, -1.185290, 1.570796, 1.834376],accel_mss,speed_ms,0,blend_radius_m)
  speed_ms = 0.005
  movel([0.263580, -0.704243, -2.808786, -1.199360, 1.570796, 1.834376],accel_mss,speed_ms,0,blend_radius_m)
  speed_ms = 0.040
  movel([0.294514, -0.677245, -2.811948, -1.223197, 1.570796, 1.865311],accel_mss,speed_ms,0,blend_radius_m)
  speed_ms = 0.005
  movel([0.294514, -0.684315, -2.818624, -1.209450, 1.570796, 1.865311],accel_mss,speed_ms,0,blend_radius_m)
  speed_ms = 0.025
  movel([0.295315, -0.680889, -2.819005, -1.212495, 1.570796, 1.866111],accel_mss,speed_ms,0,blend_radius_m)
  movel([0.296522, -0.677223, -2.819407, -1.215759, 1.570796, 1.867318],accel_mss,speed_ms,0,blend_radius_m)
  movel([0.298113, -0.673381, -2.819822, -1.219187, 1.570796, 1.868909],accel_mss,speed_ms,0,blend_radius_m)
  movel([0.300079, -0.669407, -2.820244, -1.222738, 1.570796, 1.870875],accel_mss,speed_ms,0,blend_radius_m)
  movel([0.301662, -0.666613, -2.820538, -1.225238, 1.570796, 1.872459],accel_mss,speed_ms,0,blend_radius_m)
  movel([0.303456, -0.663820, -2.820827, -1.227741, 1.570796, 1.874252],accel_mss,speed_ms,0,blend_radius_m)
  movel([0.305446, -0.661144, -2.821102, -1.230143, 1.570796, 1.876242],accel_mss,speed_ms,0,blend_radius_m)
  movel([0.307642, -0.658669, -2.821354, -1.232367, 1.570796, 1.878438],accel_mss,speed_ms,0,blend_radius_m)
  movel([0.309571, -0.656942, -2.821528, -1.233919, 1.570796, 1.880367],accel_mss,speed_ms,0,blend_radius_m)
  movel([0.311622, -0.655522, -2.821670, -1.235198, 1.570796, 1.882418],accel_mss,speed_ms,0,blend_radius_m)
  movel([0.313735, -0.654371, -2.821784, -1.236234, 1.570796, 1.884531],accel_mss,speed_ms,0,blend_radius_m)
  movel([0.315866, -0.653450, -2.821876, -1.237063, 1.570796, 1.886662],accel_mss,speed_ms,0,blend_radius_m)
  movel([0.319952, -0.652138, -2.822005, -1.238246, 1.570796, 1.890749],accel_mss,speed_ms,0,blend_radius_m)
  movel([0.323464, -0.651278, -2.822090, -1.239022, 1.570796, 1.894260],accel_mss,speed_ms,0,blend_radius_m)
  movel([0.320966, -0.652136, -2.822005, -1.238247, 1.570796, 1.891763],accel_mss,speed_ms,0,blend_radius_m)
  movel([0.318294, -0.653581, -2.821863, -1.236945, 1.570796, 1.889090],accel_mss,speed_ms,0,blend_radius_m)
  movel([0.315495, -0.655650, -2.821657, -1.235082, 1.570796, 1.886291],accel_mss,speed_ms,0,blend_radius_m)
  movel([0.312607, -0.658394, -2.821381, -1.232613, 1.570796, 1.883404],accel_mss,speed_ms,0,blend_radius_m)
  movel([0.310230, -0.661182, -2.821098, -1.230109, 1.570796, 1.881027],accel_mss,speed_ms,0,blend_radius_m)
  movel([0.308059, -0.664156, -2.820793, -1.227440, 1.570796, 1.878855],accel_mss,speed_ms,0,blend_radius_m)
  movel([0.306173, -0.667057, -2.820491, -1.224841, 1.570796, 1.876970],accel_mss,speed_ms,0,blend_radius_m)
  movel([0.304516, -0.669959, -2.820186, -1.222244, 1.570796, 1.875313],accel_mss,speed_ms,0,blend_radius_m)
  movel([0.301852, -0.675677, -2.819574, -1.217137, 1.570796, 1.872648],accel_mss,speed_ms,0,blend_radius_m)
  movel([0.300013, -0.681107, -2.818981, -1.212301, 1.570796, 1.870810],accel_mss,speed_ms,0,blend_radius_m)
  movel([0.298883, -0.686472, -2.818382, -1.207535, 1.570796, 1.869680],accel_mss,speed_ms,0,blend_radius_m)
  speed_ms = 0.005
  movel([0.298883, -0.679371, -2.811710, -1.221308, 1.570796, 1.869680],accel_mss,speed_ms,0,blend_radius_m)
  speed_ms = 0.040
  movel([0.307826, -0.665496, -2.813225, -1.233667, 1.570796, 1.878622],accel_mss,speed_ms,0,blend_radius_m)
  speed_ms = 0.005
  movel([0.307826, -0.672391, -2.819927, -1.220070, 1.570796, 1.878622],accel_mss,speed_ms,0,blend_radius_m)
  speed_ms = 0.025
  movel([0.307323, -0.673294, -2.819831, -1.219264, 1.570796, 1.878120],accel_mss,speed_ms,0,blend_radius_m)
  movel([0.306534, -0.673887, -2.819767, -1.218735, 1.570796, 1.877330],accel_mss,speed_ms,0,blend_radius_m)
  movel([0.306123, -0.673665, -2.819791, -1.218933, 1.570796, 1.876919],accel_mss,speed_ms,0,blend_radius_m)
  movel([0.306171, -0.672916, -2.819871, -1.219602, 1.570796, 1.876967],accel_mss,speed_ms,0,blend_radius_m)
  movel([0.307220, -0.670966, -2.820079, -1.221343, 1.570796, 1.878017],accel_mss,speed_ms,0,blend_radius_m)
  movel([0.307888, -0.670135, -2.820167, -1.222086, 1.570796, 1.878685],accel_mss,speed_ms,0,blend_radius_m)
  movel([0.308573, -0.669825, -2.820200, -1.222364, 1.570796, 1.879369],accel_mss,speed_ms,0,blend_radius_m)
  movel([0.308862, -0.670225, -2.820158, -1.222006, 1.570796, 1.879658],accel_mss,speed_ms,0,blend_radius_m)
  movel([0.308310, -0.671972, -2.819972, -1.220444, 1.570796, 1.879106],accel_mss,speed_ms,0,blend_radius_m)
  speed_ms = 0.005
  movel([0.308310, -0.665084, -2.813269, -1.234036, 1.570796, 1.879106],accel_mss,speed_ms,0,blend_radius_m)
  speed_ms = 0.040
  movel([0.304559, -0.685918, -2.810966, -1.215505, 1.570796, 1.875355],accel_mss,speed_ms,0,blend_radius_m)
  speed_ms = 0.005
  movel([0.304559, -0.693115, -2.817624, -1.201651, 1.570796, 1.875355],accel_mss,speed_ms,0,blend_radius_m)
  speed_ms = 0.025
  movel([0.307350, -0.689482, -2.818041, -1.204866, 1.570796, 1.878147],accel_mss,speed_ms,0,blend_radius_m)
  movel([0.309763, -0.685813, -2.818456, -1.208120, 1.570796, 1.880560],accel_mss,speed_ms,0,blend_radius_m)
  movel([0.314630, -0.678392, -2.819279, -1.214718, 1.570796, 1.885426],accel_mss,speed_ms,0,blend_radius_m)
  movel([0.318636, -0.673290, -2.819831, -1.219268, 1.570796, 1.889433],accel_mss,speed_ms,0,blend_radius_m)
  movel([0.331896, -0.658107, -2.821410, -1.232872, 1.570796, 1.902692],accel_mss,speed_ms,0,blend_radius_m)
  movel([0.334477, -0.654748, -2.821747, -1.235894, 1.570796, 1.905274],accel_mss,speed_ms,0,blend_radius_m)
  movel([0.335379, -0.653117, -2.821908, -1.237363, 1.570796, 1.906176],accel_mss,speed_ms,0,blend_radius_m)
  movel([0.335707, -0.651753, -2.822043, -1.238593, 1.570796, 1.906504],accel_mss,speed_ms,0,blend_radius_m)
  movel([0.335153, -0.650877, -2.822129, -1.239383, 1.570796, 1.905949],accel_mss,speed_ms,0,blend_radius_m)
  movel([0.333998, -0.650734, -2.822143, -1.239512, 1.570796, 1.904794],accel_mss,speed_ms,0,blend_radius_m)
  movel([0.332045, -0.650974, -2.822119, -1.239296, 1.570796, 1.902842],accel_mss,speed_ms,0,blend_radius_m)
  movel([0.330008, -0.651764, -2.822042, -1.238583, 1.570796, 1.900805],accel_mss,speed_ms,0,blend_radius_m)
  movel([0.327741, -0.653206, -2.821900, -1.237284, 1.570796, 1.898538],accel_mss,speed_ms,0,blend_radius_m)
  movel([0.325107, -0.655391, -2.821683, -1.235315, 1.570796, 1.895903],accel_mss,speed_ms,0,blend_radius_m)
  movel([0.322275, -0.658205, -2.821400, -1.232783, 1.570796, 1.893072],accel_mss,speed_ms,0,blend_radius_m)
  movel([0.319474, -0.661444, -2.821071, -1.229874, 1.570796, 1.890270],accel_mss,speed_ms,0,blend_radius_m)
  movel([0.316738, -0.664975, -2.820708, -1.226706, 1.570796, 1.887534],accel_mss,speed_ms,0,blend_radius_m)
  movel([0.314093, -0.668698, -2.820319, -1.223372, 1.570796, 1.884890],accel_mss,speed_ms,0,blend_radius_m)
  movel([0.309214, -0.676216, -2.819516, -1.216657, 1.570796, 1.880010],accel_mss,speed_ms,0,blend_radius_m)
  movel([0.305058, -0.683089, -2.818761, -1.210539, 1.570796, 1.875854],accel_mss,speed_ms,0,blend_radius_m)
  movel([0.297750, -0.695713, -2.817322, -1.199354, 1.570796, 1.868546],accel_mss,speed_ms,0,blend_radius_m)
  movel([0.295156, -0.699849, -2.816835, -1.195704, 1.570796, 1.865953],accel_mss,speed_ms,0,blend_radius_m)
  movel([0.292310, -0.703933, -2.816348, -1.192108, 1.570796, 1.863107],accel_mss,speed_ms,0,blend_radius_m)
  movel([0.289213, -0.707818, -2.815877, -1.188694, 1.570796, 1.860010],accel_mss,speed_ms,0,blend_radius_m)
  movel([0.285948, -0.711289, -2.815451, -1.185649, 1.570796, 1.856744],accel_mss,speed_ms,0,blend_radius_m)
  movel([0.282594, -0.714135, -2.815097, -1.183157, 1.570796, 1.853391],accel_mss,speed_ms,0,blend_radius_m)
  movel([0.285026, -0.713020, -2.815236, -1.184133, 1.570796, 1.855822],accel_mss,speed_ms,0,blend_radius_m)
  movel([0.287555, -0.711594, -2.815413, -1.185383, 1.570796, 1.858351],accel_mss,speed_ms,0,blend_radius_m)
  movel([0.290159, -0.709862, -2.815626, -1.186901, 1.570796, 1.860956],accel_mss,speed_ms,0,blend_radius_m)
  movel([0.292797, -0.707857, -2.815872, -1.188660, 1.570796, 1.863593],accel_mss,speed_ms,0,blend_radius_m)
  movel([0.292190, -0.710987, -2.815488, -1.185914, 1.570796, 1.862987],accel_mss,speed_ms,0,blend_radius_m)
  movel([0.291131, -0.714371, -2.815068, -1.182950, 1.570796, 1.861928],accel_mss,speed_ms,0,blend_radius_m)
  movel([0.289656, -0.717919, -2.814622, -1.179848, 1.570796, 1.860452],accel_mss,speed_ms,0,blend_radius_m)
  movel([0.287799, -0.721547, -2.814160, -1.176682, 1.570796, 1.858595],accel_mss,speed_ms,0,blend_radius_m)
  movel([0.290896, -0.717695, -2.814650, -1.180044, 1.570796, 1.861693],accel_mss,speed_ms,0,blend_radius_m)
  movel([0.293713, -0.713701, -2.815151, -1.183537, 1.570796, 1.864509],accel_mss,speed_ms,0,blend_radius_m)
  movel([0.296264, -0.709598, -2.815659, -1.187132, 1.570796, 1.867061],accel_mss,speed_ms,0,blend_radius_m)
  movel([0.298581, -0.705416, -2.816169, -1.190804, 1.570796, 1.869377],accel_mss,speed_ms,0,blend_radius_m)
  movel([0.298272, -0.707467, -2.815920, -1.189002, 1.570796, 1.869068],accel_mss,speed_ms,0,blend_radius_m)
  movel([0.297501, -0.709959, -2.815615, -1.186816, 1.570796, 1.868297],accel_mss,speed_ms,0,blend_radius_m)
  movel([0.292554, -0.721726, -2.814137, -1.176526, 1.570796, 1.863350],accel_mss,speed_ms,0,blend_radius_m)
  movel([0.291541, -0.724503, -2.813779, -1.174107, 1.570796, 1.862338],accel_mss,speed_ms,0,blend_radius_m)
  movel([0.290895, -0.726961, -2.813459, -1.171969, 1.570796, 1.861691],accel_mss,speed_ms,0,blend_radius_m)
  movel([0.292970, -0.722818, -2.813996, -1.175575, 1.570796, 1.863766],accel_mss,speed_ms,0,blend_radius_m)
  movel([0.295199, -0.718901, -2.814497, -1.178991, 1.570796, 1.865996],accel_mss,speed_ms,0,blend_radius_m)
  movel([0.300007, -0.711483, -2.815427, -1.185479, 1.570796, 1.870804],accel_mss,speed_ms,0,blend_radius_m)
  movel([0.305109, -0.704121, -2.816325, -1.191943, 1.570796, 1.875905],accel_mss,speed_ms,0,blend_radius_m)
  movel([0.310320, -0.696195, -2.817265, -1.198928, 1.570796, 1.881117],accel_mss,speed_ms,0,blend_radius_m)
  movel([0.313168, -0.691221, -2.817842, -1.203326, 1.570796, 1.883964],accel_mss,speed_ms,0,blend_radius_m)
  movel([0.314986, -0.688436, -2.818160, -1.205794, 1.570796, 1.885783],accel_mss,speed_ms,0,blend_radius_m)
  movel([0.315838, -0.687399, -2.818277, -1.206713, 1.570796, 1.886634],accel_mss,speed_ms,0,blend_radius_m)
  movel([0.316599, -0.686755, -2.818350, -1.207284, 1.570796, 1.887396],accel_mss,speed_ms,0,blend_radius_m)
  movel([0.317214, -0.686577, -2.818370, -1.207441, 1.570796, 1.888010],accel_mss,speed_ms,0,blend_radius_m)
  movel([0.317670, -0.686796, -2.818345, -1.207248, 1.570796, 1.888466],accel_mss,speed_ms,0,blend_radius_m)
  movel([0.318149, -0.688068, -2.818202, -1.206119, 1.570796, 1.888946],accel_mss,speed_ms,0,blend_radius_m)
  movel([0.318083, -0.689907, -2.817992, -1.204490, 1.570796, 1.888880],accel_mss,speed_ms,0,blend_radius_m)
  movel([0.317519, -0.691649, -2.817793, -1.202948, 1.570796, 1.888316],accel_mss,speed_ms,0,blend_radius_m)
  movel([0.320699, -0.685355, -2.818508, -1.208527, 1.570796, 1.891495],accel_mss,speed_ms,0,blend_radius_m)
  movel([0.323397, -0.679140, -2.819197, -1.214052, 1.570796, 1.894193],accel_mss,speed_ms,0,blend_radius_m)
  movel([0.325579, -0.673100, -2.819852, -1.219437, 1.570796, 1.896375],accel_mss,speed_ms,0,blend_radius_m)
  movel([0.327197, -0.667326, -2.820463, -1.224600, 1.570796, 1.897993],accel_mss,speed_ms,0,blend_radius_m)
  speed_ms = 0.005
  movel([0.327197, -0.660507, -2.813750, -1.238131, 1.570796, 1.897993],accel_mss,speed_ms,0,blend_radius_m)
  speed_ms = 0.040
  movel([0.331771, -0.660745, -2.813725, -1.237918, 1.570796, 1.902567],accel_mss,speed_ms,0,blend_radius_m)
  speed_ms = 0.005
  movel([0.331771, -0.667568, -2.820438, -1.224384, 1.570796, 1.902567],accel_mss,speed_ms,0,blend_radius_m)
  speed_ms = 0.025
  movel([0.334530, -0.667381, -2.820457, -1.224550, 1.570796, 1.905327],accel_mss,speed_ms,0,blend_radius_m)
  movel([0.335469, -0.667886, -2.820404, -1.224099, 1.570796, 1.906265],accel_mss,speed_ms,0,blend_radius_m)
  movel([0.335833, -0.669046, -2.820282, -1.223060, 1.570796, 1.906629],accel_mss,speed_ms,0,blend_radius_m)
  movel([0.335591, -0.670536, -2.820125, -1.221728, 1.570796, 1.906388],accel_mss,speed_ms,0,blend_radius_m)
  movel([0.326578, -0.697817, -2.817075, -1.197497, 1.570796, 1.897374],accel_mss,speed_ms,0,blend_radius_m)
  movel([0.325852, -0.699779, -2.816844, -1.195766, 1.570796, 1.896648],accel_mss,speed_ms,0,blend_radius_m)
  movel([0.324885, -0.701813, -2.816602, -1.193975, 1.570796, 1.895681],accel_mss,speed_ms,0,blend_radius_m)
  movel([0.323657, -0.703672, -2.816379, -1.192338, 1.570796, 1.894453],accel_mss,speed_ms,0,blend_radius_m)
  movel([0.322169, -0.705103, -2.816207, -1.191080, 1.570796, 1.892965],accel_mss,speed_ms,0,blend_radius_m)
  movel([0.320845, -0.705716, -2.816132, -1.190541, 1.570796, 1.891642],accel_mss,speed_ms,0,blend_radius_m)
  movel([0.318504, -0.706023, -2.816095, -1.190270, 1.570796, 1.889300],accel_mss,speed_ms,0,blend_radius_m)
  movel([0.317175, -0.706703, -2.816013, -1.189673, 1.570796, 1.887972],accel_mss,speed_ms,0,blend_radius_m)
  movel([0.315504, -0.708415, -2.815804, -1.188170, 1.570796, 1.886301],accel_mss,speed_ms,0,blend_radius_m)
  movel([0.313959, -0.710461, -2.815553, -1.186375, 1.570796, 1.884756],accel_mss,speed_ms,0,blend_radius_m)
  movel([0.312038, -0.712771, -2.815267, -1.184351, 1.570796, 1.882835],accel_mss,speed_ms,0,blend_radius_m)
  movel([0.309999, -0.714812, -2.815013, -1.182564, 1.570796, 1.880795],accel_mss,speed_ms,0,blend_radius_m)
  movel([0.307917, -0.716539, -2.814796, -1.181054, 1.570796, 1.878713],accel_mss,speed_ms,0,blend_radius_m)
  movel([0.305858, -0.717914, -2.814622, -1.179853, 1.570796, 1.876655],accel_mss,speed_ms,0,blend_radius_m)
  movel([0.303892, -0.718900, -2.814497, -1.178991, 1.570796, 1.874689],accel_mss,speed_ms,0,blend_radius_m)
  movel([0.302101, -0.719445, -2.814428, -1.178516, 1.570796, 1.872898],accel_mss,speed_ms,0,blend_radius_m)
  movel([0.300546, -0.719525, -2.814418, -1.178446, 1.570796, 1.871343],accel_mss,speed_ms,0,blend_radius_m)
  movel([0.299304, -0.719079, -2.814475, -1.178836, 1.570796, 1.870100],accel_mss,speed_ms,0,blend_radius_m)
  speed_ms = 0.005
  movel([0.299304, -0.711522, -2.807878, -1.192989, 1.570796, 1.870100],accel_mss,speed_ms,0,blend_radius_m)
  speed_ms = 0.040
  movel([0.281741, -0.738260, -2.804338, -1.169791, 1.570796, 1.852537],accel_mss,speed_ms,0,blend_radius_m)
  speed_ms = 0.005
  movel([0.281741, -0.746167, -2.810866, -1.155356, 1.570796, 1.852537],accel_mss,speed_ms,0,blend_radius_m)
  speed_ms = 0.025
  movel([0.278055, -0.769343, -2.807506, -1.135540, 1.570796, 1.848852],accel_mss,speed_ms,0,blend_radius_m)
  movel([0.277347, -0.772302, -2.807059, -1.133028, 1.570796, 1.848143],accel_mss,speed_ms,0,blend_radius_m)
  movel([0.276648, -0.773846, -2.806823, -1.131719, 1.570796, 1.847444],accel_mss,speed_ms,0,blend_radius_m)
  movel([0.275612, -0.775338, -2.806595, -1.130456, 1.570796, 1.846408],accel_mss,speed_ms,0,blend_radius_m)
  movel([0.272899, -0.778154, -2.806161, -1.128074, 1.570796, 1.843695],accel_mss,speed_ms,0,blend_radius_m)
  movel([0.271996, -0.779823, -2.805902, -1.126665, 1.570796, 1.842792],accel_mss,speed_ms,0,blend_radius_m)
  movel([0.271579, -0.781403, -2.805655, -1.125331, 1.570796, 1.842375],accel_mss,speed_ms,0,blend_radius_m)
  movel([0.271570, -0.783618, -2.805307, -1.123464, 1.570796, 1.842366],accel_mss,speed_ms,0,blend_radius_m)
  movel([0.272150, -0.785418, -2.805023, -1.121948, 1.570796, 1.842946],accel_mss,speed_ms,0,blend_radius_m)
  movel([0.273739, -0.788498, -2.804532, -1.119358, 1.570796, 1.844535],accel_mss,speed_ms,0,blend_radius_m)
  movel([0.274278, -0.791015, -2.804128, -1.117246, 1.570796, 1.845075],accel_mss,speed_ms,0,blend_radius_m)
  movel([0.274468, -0.795049, -2.803473, -1.113867, 1.570796, 1.845264],accel_mss,speed_ms,0,blend_radius_m)
  movel([0.274204, -0.797087, -2.803139, -1.112163, 1.570796, 1.845000],accel_mss,speed_ms,0,blend_radius_m)
  movel([0.273576, -0.798865, -2.802846, -1.110678, 1.570796, 1.844372],accel_mss,speed_ms,0,blend_radius_m)
  movel([0.273096, -0.799582, -2.802727, -1.110079, 1.570796, 1.843892],accel_mss,speed_ms,0,blend_radius_m)
  movel([0.272493, -0.800157, -2.802632, -1.109600, 1.570796, 1.843289],accel_mss,speed_ms,0,blend_radius_m)
  movel([0.271753, -0.800561, -2.802565, -1.109263, 1.570796, 1.842549],accel_mss,speed_ms,0,blend_radius_m)
  movel([0.270866, -0.800762, -2.802532, -1.109096, 1.570796, 1.841663],accel_mss,speed_ms,0,blend_radius_m)
  movel([0.270373, -0.802611, -2.802223, -1.107555, 1.570796, 1.841169],accel_mss,speed_ms,0,blend_radius_m)
  movel([0.270264, -0.804477, -2.801910, -1.106002, 1.570796, 1.841060],accel_mss,speed_ms,0,blend_radius_m)
  movel([0.270864, -0.808104, -2.801297, -1.102988, 1.570796, 1.841661],accel_mss,speed_ms,0,blend_radius_m)
  movel([0.272032, -0.811284, -2.800753, -1.100352, 1.570796, 1.842829],accel_mss,speed_ms,0,blend_radius_m)
  movel([0.273153, -0.813648, -2.800346, -1.098395, 1.570796, 1.843949],accel_mss,speed_ms,0,blend_radius_m)
  movel([0.274846, -0.815814, -2.799970, -1.096605, 1.570796, 1.845642],accel_mss,speed_ms,0,blend_radius_m)
  movel([0.276926, -0.817721, -2.799637, -1.095031, 1.570796, 1.847722],accel_mss,speed_ms,0,blend_radius_m)
  movel([0.278568, -0.820032, -2.799231, -1.093126, 1.570796, 1.849364],accel_mss,speed_ms,0,blend_radius_m)
  movel([0.278969, -0.821535, -2.798965, -1.091888, 1.570796, 1.849766],accel_mss,speed_ms,0,blend_radius_m)
  movel([0.278953, -0.823381, -2.798638, -1.090371, 1.570796, 1.849750],accel_mss,speed_ms,0,blend_radius_m)
  movel([0.278680, -0.824495, -2.798439, -1.089456, 1.570796, 1.849477],accel_mss,speed_ms,0,blend_radius_m)
  movel([0.278145, -0.825700, -2.798223, -1.088466, 1.570796, 1.848941],accel_mss,speed_ms,0,blend_radius_m)
  movel([0.277410, -0.826747, -2.798035, -1.087607, 1.570796, 1.848207],accel_mss,speed_ms,0,blend_radius_m)
  movel([0.276534, -0.827400, -2.797917, -1.087072, 1.570796, 1.847330],accel_mss,speed_ms,0,blend_radius_m)
  movel([0.275921, -0.827455, -2.797907, -1.087027, 1.570796, 1.846718],accel_mss,speed_ms,0,blend_radius_m)
  movel([0.275468, -0.827227, -2.797948, -1.087213, 1.570796, 1.846264],accel_mss,speed_ms,0,blend_radius_m)
  movel([0.271858, -0.824094, -2.798510, -1.089785, 1.570796, 1.842655],accel_mss,speed_ms,0,blend_radius_m)
  movel([0.270330, -0.822188, -2.798850, -1.091352, 1.570796, 1.841127],accel_mss,speed_ms,0,blend_radius_m)
  movel([0.269001, -0.820052, -2.799228, -1.093109, 1.570796, 1.839798],accel_mss,speed_ms,0,blend_radius_m)
  movel([0.268223, -0.821276, -2.799011, -1.092101, 1.570796, 1.839019],accel_mss,speed_ms,0,blend_radius_m)
  movel([0.267662, -0.822501, -2.798794, -1.091094, 1.570796, 1.838458],accel_mss,speed_ms,0,blend_radius_m)
  movel([0.267117, -0.824921, -2.798363, -1.089105, 1.570796, 1.837913],accel_mss,speed_ms,0,blend_radius_m)
  movel([0.267194, -0.827260, -2.797943, -1.087187, 1.570796, 1.837990],accel_mss,speed_ms,0,blend_radius_m)
  movel([0.267740, -0.829458, -2.797545, -1.085386, 1.570796, 1.838537],accel_mss,speed_ms,0,blend_radius_m)
  movel([0.269558, -0.833265, -2.796851, -1.082273, 1.570796, 1.840354],accel_mss,speed_ms,0,blend_radius_m)
  movel([0.271292, -0.835911, -2.796363, -1.080115, 1.570796, 1.842088],accel_mss,speed_ms,0,blend_radius_m)
  movel([0.271782, -0.837044, -2.796153, -1.079191, 1.570796, 1.842578],accel_mss,speed_ms,0,blend_radius_m)
  movel([0.271770, -0.837787, -2.796016, -1.078587, 1.570796, 1.842567],accel_mss,speed_ms,0,blend_radius_m)
  movel([0.271447, -0.838685, -2.795848, -1.077856, 1.570796, 1.842243],accel_mss,speed_ms,0,blend_radius_m)
  movel([0.270811, -0.839658, -2.795667, -1.077064, 1.570796, 1.841608],accel_mss,speed_ms,0,blend_radius_m)
  movel([0.270166, -0.840263, -2.795554, -1.076573, 1.570796, 1.840962],accel_mss,speed_ms,0,blend_radius_m)
  movel([0.268900, -0.840739, -2.795464, -1.076186, 1.570796, 1.839696],accel_mss,speed_ms,0,blend_radius_m)
  movel([0.267192, -0.841164, -2.795384, -1.075840, 1.570796, 1.837988],accel_mss,speed_ms,0,blend_radius_m)
  movel([0.266720, -0.841632, -2.795297, -1.075461, 1.570796, 1.837517],accel_mss,speed_ms,0,blend_radius_m)
  movel([0.266266, -0.842481, -2.795137, -1.074771, 1.570796, 1.837062],accel_mss,speed_ms,0,blend_radius_m)
  movel([0.266043, -0.843369, -2.794969, -1.074050, 1.570796, 1.836840],accel_mss,speed_ms,0,blend_radius_m)
  movel([0.266116, -0.845145, -2.794633, -1.072611, 1.570796, 1.836912],accel_mss,speed_ms,0,blend_radius_m)
  movel([0.266945, -0.847921, -2.794103, -1.070365, 1.570796, 1.837741],accel_mss,speed_ms,0,blend_radius_m)
  movel([0.269138, -0.853386, -2.793048, -1.065955, 1.570796, 1.839934],accel_mss,speed_ms,0,blend_radius_m)
  movel([0.271450, -0.858701, -2.792006, -1.061683, 1.570796, 1.842246],accel_mss,speed_ms,0,blend_radius_m)
  movel([0.271715, -0.859953, -2.791758, -1.060678, 1.570796, 1.842512],accel_mss,speed_ms,0,blend_radius_m)
  movel([0.271667, -0.861446, -2.791461, -1.059482, 1.570796, 1.842463],accel_mss,speed_ms,0,blend_radius_m)
  movel([0.271156, -0.863037, -2.791143, -1.058209, 1.570796, 1.841952],accel_mss,speed_ms,0,blend_radius_m)
  movel([0.270689, -0.863819, -2.790987, -1.057583, 1.570796, 1.841485],accel_mss,speed_ms,0,blend_radius_m)
  movel([0.269378, -0.865146, -2.790720, -1.056523, 1.570796, 1.840175],accel_mss,speed_ms,0,blend_radius_m)
  movel([0.268742, -0.865509, -2.790647, -1.056233, 1.570796, 1.839539],accel_mss,speed_ms,0,blend_radius_m)
  movel([0.267584, -0.865702, -2.790608, -1.056079, 1.570796, 1.838380],accel_mss,speed_ms,0,blend_radius_m)
  movel([0.266607, -0.865378, -2.790673, -1.056338, 1.570796, 1.837403],accel_mss,speed_ms,0,blend_radius_m)
  movel([0.265848, -0.864746, -2.790800, -1.056843, 1.570796, 1.836644],accel_mss,speed_ms,0,blend_radius_m)
  movel([0.262076, -0.860186, -2.791711, -1.060492, 1.570796, 1.832873],accel_mss,speed_ms,0,blend_radius_m)
  movel([0.258644, -0.855210, -2.792692, -1.064487, 1.570796, 1.829441],accel_mss,speed_ms,0,blend_radius_m)
  movel([0.255575, -0.849810, -2.793740, -1.068839, 1.570796, 1.826371],accel_mss,speed_ms,0,blend_radius_m)
  movel([0.252877, -0.843987, -2.794852, -1.073549, 1.570796, 1.823673],accel_mss,speed_ms,0,blend_radius_m)
  movel([0.252039, -0.841663, -2.795291, -1.075436, 1.570796, 1.822835],accel_mss,speed_ms,0,blend_radius_m)
  movel([0.251666, -0.838933, -2.795802, -1.077654, 1.570796, 1.822462],accel_mss,speed_ms,0,blend_radius_m)
  movel([0.251810, -0.837040, -2.796154, -1.079195, 1.570796, 1.822606],accel_mss,speed_ms,0,blend_radius_m)
  movel([0.252185, -0.835001, -2.796531, -1.080857, 1.570796, 1.822981],accel_mss,speed_ms,0,blend_radius_m)
  movel([0.253320, -0.830686, -2.797322, -1.084381, 1.570796, 1.824117],accel_mss,speed_ms,0,blend_radius_m)
  movel([0.258739, -0.814486, -2.800201, -1.097702, 1.570796, 1.829535],accel_mss,speed_ms,0,blend_radius_m)
  movel([0.259950, -0.810007, -2.800972, -1.101410, 1.570796, 1.830746],accel_mss,speed_ms,0,blend_radius_m)
  movel([0.260608, -0.806159, -2.801627, -1.104603, 1.570796, 1.831404],accel_mss,speed_ms,0,blend_radius_m)
  movel([0.260657, -0.804598, -2.801890, -1.105901, 1.570796, 1.831453],accel_mss,speed_ms,0,blend_radius_m)
  movel([0.260469, -0.803355, -2.802099, -1.106936, 1.570796, 1.831265],accel_mss,speed_ms,0,blend_radius_m)
  movel([0.260019, -0.802474, -2.802246, -1.107669, 1.570796, 1.830816],accel_mss,speed_ms,0,blend_radius_m)
  movel([0.259280, -0.802008, -2.802324, -1.108057, 1.570796, 1.830076],accel_mss,speed_ms,0,blend_radius_m)
  movel([0.257564, -0.801881, -2.802345, -1.108163, 1.570796, 1.828361],accel_mss,speed_ms,0,blend_radius_m)
  movel([0.256825, -0.801681, -2.802379, -1.108330, 1.570796, 1.827621],accel_mss,speed_ms,0,blend_radius_m)
  movel([0.256410, -0.801087, -2.802477, -1.108824, 1.570796, 1.827206],accel_mss,speed_ms,0,blend_radius_m)
  movel([0.256635, -0.799469, -2.802746, -1.110174, 1.570796, 1.827431],accel_mss,speed_ms,0,blend_radius_m)
  movel([0.257472, -0.797499, -2.803071, -1.111818, 1.570796, 1.828269],accel_mss,speed_ms,0,blend_radius_m)
  movel([0.260367, -0.791124, -2.804110, -1.117155, 1.570796, 1.831164],accel_mss,speed_ms,0,blend_radius_m)
  movel([0.262974, -0.784821, -2.805117, -1.122451, 1.570796, 1.833770],accel_mss,speed_ms,0,blend_radius_m)
  movel([0.265331, -0.778565, -2.806097, -1.127727, 1.570796, 1.836127],accel_mss,speed_ms,0,blend_radius_m)
  movel([0.267477, -0.772341, -2.807053, -1.132996, 1.570796, 1.838273],accel_mss,speed_ms,0,blend_radius_m)
  movel([0.271335, -0.759911, -2.808905, -1.143573, 1.570796, 1.842131],accel_mss,speed_ms,0,blend_radius_m)
  movel([0.274904, -0.747355, -2.810700, -1.154334, 1.570796, 1.845701],accel_mss,speed_ms,0,blend_radius_m)
  speed_ms = 0.005
  movel([0.274904, -0.739433, -2.804175, -1.168781, 1.570796, 1.845701],accel_mss,speed_ms,0,blend_radius_m)
  speed_ms = 0.040
  movel([0.261432, -0.771781, -2.799423, -1.141185, 1.570796, 1.832228],accel_mss,speed_ms,0,blend_radius_m)
  speed_ms = 0.005
  movel([0.261432, -0.780092, -2.805860, -1.126437, 1.570796, 1.832228],accel_mss,speed_ms,0,blend_radius_m)
  speed_ms = 0.025
  movel([0.254948, -0.788762, -2.804490, -1.119137, 1.570796, 1.825745],accel_mss,speed_ms,0,blend_radius_m)
  movel([0.248348, -0.797178, -2.803124, -1.112087, 1.570796, 1.819145],accel_mss,speed_ms,0,blend_radius_m)
  movel([0.241644, -0.805338, -2.801765, -1.105286, 1.570796, 1.812440],accel_mss,speed_ms,0,blend_radius_m)
  movel([0.234856, -0.813215, -2.800421, -1.098753, 1.570796, 1.805652],accel_mss,speed_ms,0,blend_radius_m)
  movel([0.240164, -0.805142, -2.801798, -1.105449, 1.570796, 1.810961],accel_mss,speed_ms,0,blend_radius_m)
  movel([0.245154, -0.796888, -2.803172, -1.112329, 1.570796, 1.815950],accel_mss,speed_ms,0,blend_radius_m)
  movel([0.249787, -0.788509, -2.804530, -1.119350, 1.570796, 1.820583],accel_mss,speed_ms,0,blend_radius_m)
  movel([0.254028, -0.780060, -2.805865, -1.126465, 1.570796, 1.824825],accel_mss,speed_ms,0,blend_radius_m)
  movel([0.248584, -0.787180, -2.804743, -1.120467, 1.570796, 1.819380],accel_mss,speed_ms,0,blend_radius_m)
  movel([0.243053, -0.794107, -2.803627, -1.114656, 1.570796, 1.813849],accel_mss,speed_ms,0,blend_radius_m)
  movel([0.237436, -0.800841, -2.802518, -1.109030, 1.570796, 1.808232],accel_mss,speed_ms,0,blend_radius_m)
  movel([0.231748, -0.807361, -2.801423, -1.103605, 1.570796, 1.802544],accel_mss,speed_ms,0,blend_radius_m)
  movel([0.225400, -0.814446, -2.800208, -1.097735, 1.570796, 1.796196],accel_mss,speed_ms,0,blend_radius_m)
  movel([0.219321, -0.821682, -2.798939, -1.091768, 1.570796, 1.790117],accel_mss,speed_ms,0,blend_radius_m)
  movel([0.216506, -0.825477, -2.798263, -1.088649, 1.570796, 1.787302],accel_mss,speed_ms,0,blend_radius_m)
  movel([0.213960, -0.829363, -2.797562, -1.085463, 1.570796, 1.784756],accel_mss,speed_ms,0,blend_radius_m)
  movel([0.211819, -0.833252, -2.796853, -1.082284, 1.570796, 1.782615],accel_mss,speed_ms,0,blend_radius_m)
  movel([0.210196, -0.837054, -2.796152, -1.079184, 1.570796, 1.780992],accel_mss,speed_ms,0,blend_radius_m)
  movel([0.211400, -0.832627, -2.796968, -1.082795, 1.570796, 1.782197],accel_mss,speed_ms,0,blend_radius_m)
  movel([0.212956, -0.827934, -2.797821, -1.086634, 1.570796, 1.783752],accel_mss,speed_ms,0,blend_radius_m)
  movel([0.214839, -0.823035, -2.798699, -1.090655, 1.570796, 1.785635],accel_mss,speed_ms,0,blend_radius_m)
  movel([0.217020, -0.817988, -2.799590, -1.094810, 1.570796, 1.787816],accel_mss,speed_ms,0,blend_radius_m)
  movel([0.219468, -0.812858, -2.800482, -1.099048, 1.570796, 1.790265],accel_mss,speed_ms,0,blend_radius_m)
  movel([0.222158, -0.807705, -2.801365, -1.103319, 1.570796, 1.792954],accel_mss,speed_ms,0,blend_radius_m)
  movel([0.225056, -0.802598, -2.802225, -1.107566, 1.570796, 1.795852],accel_mss,speed_ms,0,blend_radius_m)
  movel([0.228128, -0.797608, -2.803053, -1.111728, 1.570796, 1.798924],accel_mss,speed_ms,0,blend_radius_m)
  movel([0.222602, -0.805419, -2.801752, -1.105219, 1.570796, 1.793398],accel_mss,speed_ms,0,blend_radius_m)
  movel([0.217407, -0.813235, -2.800417, -1.098736, 1.570796, 1.788203],accel_mss,speed_ms,0,blend_radius_m)
  movel([0.212522, -0.821034, -2.799054, -1.092301, 1.570796, 1.783318],accel_mss,speed_ms,0,blend_radius_m)
  movel([0.207928, -0.828790, -2.797666, -1.085932, 1.570796, 1.778724],accel_mss,speed_ms,0,blend_radius_m)
  movel([0.203609, -0.836476, -2.796259, -1.079654, 1.570796, 1.774406],accel_mss,speed_ms,0,blend_radius_m)
  movel([0.199541, -0.844073, -2.794836, -1.073480, 1.570796, 1.770338],accel_mss,speed_ms,0,blend_radius_m)
  movel([0.192077, -0.858910, -2.791964, -1.061515, 1.570796, 1.762873],accel_mss,speed_ms,0,blend_radius_m)
  movel([0.194129, -0.853899, -2.792948, -1.065542, 1.570796, 1.764926],accel_mss,speed_ms,0,blend_radius_m)
  movel([0.195772, -0.848649, -2.793963, -1.069777, 1.570796, 1.766568],accel_mss,speed_ms,0,blend_radius_m)
  movel([0.198677, -0.838450, -2.795892, -1.078047, 1.570796, 1.769474],accel_mss,speed_ms,0,blend_radius_m)
  movel([0.200321, -0.833793, -2.796754, -1.081842, 1.570796, 1.771117],accel_mss,speed_ms,0,blend_radius_m)
  movel([0.202086, -0.829515, -2.797535, -1.085339, 1.570796, 1.772882],accel_mss,speed_ms,0,blend_radius_m)
  movel([0.206386, -0.820504, -2.799148, -1.092737, 1.570796, 1.777183],accel_mss,speed_ms,0,blend_radius_m)
  movel([0.205471, -0.821821, -2.798915, -1.091653, 1.570796, 1.776267],accel_mss,speed_ms,0,blend_radius_m)
  movel([0.203922, -0.823541, -2.798609, -1.090239, 1.570796, 1.774718],accel_mss,speed_ms,0,blend_radius_m)
  movel([0.195262, -0.831821, -2.797115, -1.083453, 1.570796, 1.766058],accel_mss,speed_ms,0,blend_radius_m)
  movel([0.192150, -0.834965, -2.796538, -1.080886, 1.570796, 1.762947],accel_mss,speed_ms,0,blend_radius_m)
  movel([0.188692, -0.839395, -2.795716, -1.077278, 1.570796, 1.759489],accel_mss,speed_ms,0,blend_radius_m)
  movel([0.185491, -0.844085, -2.794834, -1.073470, 1.570796, 1.756287],accel_mss,speed_ms,0,blend_radius_m)
  movel([0.179730, -0.853510, -2.793024, -1.065855, 1.570796, 1.750526],accel_mss,speed_ms,0,blend_radius_m)
  movel([0.181985, -0.848632, -2.793967, -1.069791, 1.570796, 1.752782],accel_mss,speed_ms,0,blend_radius_m)
  movel([0.183935, -0.843771, -2.794893, -1.073725, 1.570796, 1.754732],accel_mss,speed_ms,0,blend_radius_m)
  movel([0.187766, -0.833971, -2.796721, -1.081697, 1.570796, 1.758562],accel_mss,speed_ms,0,blend_radius_m)
  movel([0.190156, -0.828765, -2.797671, -1.085954, 1.570796, 1.760953],accel_mss,speed_ms,0,blend_radius_m)
  movel([0.192896, -0.823448, -2.798626, -1.090316, 1.570796, 1.763693],accel_mss,speed_ms,0,blend_radius_m)
  movel([0.199179, -0.812542, -2.800537, -1.099310, 1.570796, 1.769975],accel_mss,speed_ms,0,blend_radius_m)
  movel([0.212906, -0.790485, -2.804213, -1.117691, 1.570796, 1.783702],accel_mss,speed_ms,0,blend_radius_m)
  movel([0.207618, -0.794989, -2.803483, -1.113917, 1.570796, 1.778414],accel_mss,speed_ms,0,blend_radius_m)
  movel([0.202419, -0.799803, -2.802691, -1.109895, 1.570796, 1.773215],accel_mss,speed_ms,0,blend_radius_m)
  movel([0.197333, -0.804883, -2.801842, -1.105664, 1.570796, 1.768130],accel_mss,speed_ms,0,blend_radius_m)
  movel([0.192402, -0.810187, -2.800941, -1.101260, 1.570796, 1.763198],accel_mss,speed_ms,0,blend_radius_m)
  movel([0.187658, -0.815677, -2.799994, -1.096718, 1.570796, 1.758454],accel_mss,speed_ms,0,blend_radius_m)
  movel([0.183125, -0.821318, -2.799004, -1.092067, 1.570796, 1.753921],accel_mss,speed_ms,0,blend_radius_m)
  movel([0.178832, -0.827068, -2.797977, -1.087344, 1.570796, 1.749628],accel_mss,speed_ms,0,blend_radius_m)
  movel([0.174808, -0.832897, -2.796918, -1.082574, 1.570796, 1.745604],accel_mss,speed_ms,0,blend_radius_m)
  movel([0.175871, -0.831123, -2.797242, -1.084024, 1.570796, 1.746668],accel_mss,speed_ms,0,blend_radius_m)
  movel([0.176866, -0.829156, -2.797600, -1.085633, 1.570796, 1.747662],accel_mss,speed_ms,0,blend_radius_m)
  movel([0.178700, -0.824880, -2.798370, -1.089139, 1.570796, 1.749496],accel_mss,speed_ms,0,blend_radius_m)
  movel([0.182052, -0.816663, -2.799822, -1.095904, 1.570796, 1.752849],accel_mss,speed_ms,0,blend_radius_m)
  movel([0.185570, -0.809472, -2.801064, -1.101853, 1.570796, 1.756367],accel_mss,speed_ms,0,blend_radius_m)
  movel([0.189353, -0.802229, -2.802287, -1.107873, 1.570796, 1.760150],accel_mss,speed_ms,0,blend_radius_m)
  movel([0.193392, -0.794935, -2.803492, -1.113962, 1.570796, 1.764188],accel_mss,speed_ms,0,blend_radius_m)
  movel([0.197671, -0.787593, -2.804677, -1.120119, 1.570796, 1.768468],accel_mss,speed_ms,0,blend_radius_m)
  movel([0.202185, -0.780190, -2.805844, -1.126355, 1.570796, 1.772981],accel_mss,speed_ms,0,blend_radius_m)
  movel([0.206927, -0.772732, -2.806993, -1.132664, 1.570796, 1.777723],accel_mss,speed_ms,0,blend_radius_m)
  movel([0.217047, -0.757615, -2.809239, -1.145536, 1.570796, 1.787844],accel_mss,speed_ms,0,blend_radius_m)
  movel([0.212834, -0.762359, -2.808546, -1.141484, 1.570796, 1.783630],accel_mss,speed_ms,0,blend_radius_m)
  movel([0.199928, -0.775754, -2.806531, -1.130104, 1.570796, 1.770724],accel_mss,speed_ms,0,blend_radius_m)
  movel([0.195714, -0.780307, -2.805826, -1.126256, 1.570796, 1.766510],accel_mss,speed_ms,0,blend_radius_m)
  movel([0.191666, -0.785043, -2.805082, -1.122264, 1.570796, 1.762463],accel_mss,speed_ms,0,blend_radius_m)
  movel([0.187933, -0.789942, -2.804301, -1.118146, 1.570796, 1.758729],accel_mss,speed_ms,0,blend_radius_m)
  movel([0.184647, -0.795000, -2.803481, -1.113908, 1.570796, 1.755443],accel_mss,speed_ms,0,blend_radius_m)
  movel([0.189107, -0.786707, -2.804818, -1.120864, 1.570796, 1.759904],accel_mss,speed_ms,0,blend_radius_m)
  movel([0.193566, -0.778056, -2.806176, -1.128157, 1.570796, 1.764363],accel_mss,speed_ms,0,blend_radius_m)
  movel([0.198297, -0.769349, -2.807505, -1.135535, 1.570796, 1.769093],accel_mss,speed_ms,0,blend_radius_m)
  movel([0.200846, -0.765079, -2.808144, -1.139166, 1.570796, 1.771643],accel_mss,speed_ms,0,blend_radius_m)
  movel([0.203569, -0.760920, -2.808757, -1.142712, 1.570796, 1.774365],accel_mss,speed_ms,0,blend_radius_m)
  movel([0.213662, -0.746902, -2.810764, -1.154724, 1.570796, 1.784458],accel_mss,speed_ms,0,blend_radius_m)
  movel([0.224121, -0.732719, -2.812700, -1.166971, 1.570796, 1.794917],accel_mss,speed_ms,0,blend_radius_m)
  movel([0.216555, -0.740130, -2.811700, -1.160560, 1.570796, 1.787351],accel_mss,speed_ms,0,blend_radius_m)
  movel([0.209738, -0.747489, -2.810681, -1.154219, 1.570796, 1.780535],accel_mss,speed_ms,0,blend_radius_m)
  movel([0.203245, -0.755289, -2.809574, -1.147526, 1.570796, 1.774041],accel_mss,speed_ms,0,blend_radius_m)
  movel([0.196669, -0.763988, -2.808305, -1.140096, 1.570796, 1.767465],accel_mss,speed_ms,0,blend_radius_m)
  movel([0.199815, -0.759356, -2.808985, -1.144047, 1.570796, 1.770611],accel_mss,speed_ms,0,blend_radius_m)
  movel([0.202657, -0.754651, -2.809666, -1.148072, 1.570796, 1.773453],accel_mss,speed_ms,0,blend_radius_m)
  movel([0.213090, -0.735308, -2.812353, -1.164728, 1.570796, 1.783886],accel_mss,speed_ms,0,blend_radius_m)
  movel([0.215992, -0.730398, -2.813008, -1.168983, 1.570796, 1.786788],accel_mss,speed_ms,0,blend_radius_m)
  movel([0.219234, -0.725477, -2.813653, -1.173260, 1.570796, 1.790031],accel_mss,speed_ms,0,blend_radius_m)
  movel([0.223935, -0.719165, -2.814464, -1.178761, 1.570796, 1.794731],accel_mss,speed_ms,0,blend_radius_m)
  movel([0.228034, -0.714530, -2.815048, -1.182811, 1.570796, 1.798830],accel_mss,speed_ms,0,blend_radius_m)
  movel([0.228958, -0.713224, -2.815211, -1.183954, 1.570796, 1.799754],accel_mss,speed_ms,0,blend_radius_m)
  movel([0.229281, -0.712119, -2.815348, -1.184922, 1.570796, 1.800078],accel_mss,speed_ms,0,blend_radius_m)
  movel([0.228746, -0.711887, -2.815377, -1.185125, 1.570796, 1.799542],accel_mss,speed_ms,0,blend_radius_m)
  movel([0.227577, -0.712329, -2.815322, -1.184738, 1.570796, 1.798373],accel_mss,speed_ms,0,blend_radius_m)
  movel([0.226000, -0.713253, -2.815207, -1.183929, 1.570796, 1.796796],accel_mss,speed_ms,0,blend_radius_m)
  movel([0.222512, -0.715717, -2.814899, -1.181773, 1.570796, 1.793308],accel_mss,speed_ms,0,blend_radius_m)
  movel([0.220069, -0.717685, -2.814651, -1.180053, 1.570796, 1.790865],accel_mss,speed_ms,0,blend_radius_m)
  movel([0.223947, -0.711964, -2.815367, -1.185058, 1.570796, 1.794743],accel_mss,speed_ms,0,blend_radius_m)
  movel([0.228482, -0.706191, -2.816075, -1.190124, 1.570796, 1.799278],accel_mss,speed_ms,0,blend_radius_m)
  movel([0.237978, -0.695251, -2.817376, -1.199763, 1.570796, 1.808774],accel_mss,speed_ms,0,blend_radius_m)
  speed_ms = 0.005
  movel([0.237978, -0.688023, -2.810723, -1.213642, 1.570796, 1.808774],accel_mss,speed_ms,0,blend_radius_m)
  speed_ms = 0.040
  movel([0.220547, -0.698392, -2.809498, -1.204499, 1.570796, 1.791343],accel_mss,speed_ms,0,blend_radius_m)
  speed_ms = 0.005
  movel([0.220547, -0.705767, -2.816126, -1.190496, 1.570796, 1.791343],accel_mss,speed_ms,0,blend_radius_m)
  speed_ms = 0.025
  movel([0.219117, -0.704356, -2.816297, -1.191736, 1.570796, 1.789913],accel_mss,speed_ms,0,blend_radius_m)
  movel([0.217209, -0.703678, -2.816378, -1.192333, 1.570796, 1.788005],accel_mss,speed_ms,0,blend_radius_m)
  movel([0.214903, -0.703651, -2.816381, -1.192357, 1.570796, 1.785699],accel_mss,speed_ms,0,blend_radius_m)
  movel([0.212279, -0.704187, -2.816317, -1.191885, 1.570796, 1.783076],accel_mss,speed_ms,0,blend_radius_m)
  movel([0.209410, -0.705216, -2.816193, -1.190980, 1.570796, 1.780207],accel_mss,speed_ms,0,blend_radius_m)
  movel([0.206382, -0.706649, -2.816019, -1.189721, 1.570796, 1.777179],accel_mss,speed_ms,0,blend_radius_m)
  movel([0.200145, -0.710390, -2.815561, -1.186437, 1.570796, 1.770941],accel_mss,speed_ms,0,blend_radius_m)
  speed_ms = 0.005
  movel([0.200145, -0.702952, -2.808944, -1.200493, 1.570796, 1.770941],accel_mss,speed_ms,0,blend_radius_m)
  speed_ms = 0.040
  movel([0.225931, -0.680542, -2.811578, -1.220269, 1.570796, 1.796727],accel_mss,speed_ms,0,blend_radius_m)
  speed_ms = 0.005
  movel([0.225931, -0.687661, -2.818248, -1.206480, 1.570796, 1.796727],accel_mss,speed_ms,0,blend_radius_m)
  speed_ms = 0.025
  movel([0.225055, -0.683915, -2.818669, -1.209805, 1.570796, 1.795851],accel_mss,speed_ms,0,blend_radius_m)
  movel([0.223901, -0.680589, -2.819038, -1.212762, 1.570796, 1.794697],accel_mss,speed_ms,0,blend_radius_m)
  movel([0.222358, -0.677842, -2.819339, -1.215208, 1.570796, 1.793155],accel_mss,speed_ms,0,blend_radius_m)
  movel([0.220313, -0.675828, -2.819558, -1.217003, 1.570796, 1.791109],accel_mss,speed_ms,0,blend_radius_m)
  movel([0.217651, -0.674726, -2.819677, -1.217986, 1.570796, 1.788447],accel_mss,speed_ms,0,blend_radius_m)
  movel([0.214276, -0.674669, -2.819683, -1.218037, 1.570796, 1.785072],accel_mss,speed_ms,0,blend_radius_m)
  movel([0.210076, -0.675837, -2.819557, -1.216995, 1.570796, 1.780872],accel_mss,speed_ms,0,blend_radius_m)
  movel([0.207638, -0.676922, -2.819439, -1.216028, 1.570796, 1.778434],accel_mss,speed_ms,0,blend_radius_m)
  movel([0.204957, -0.678369, -2.819282, -1.214739, 1.570796, 1.775753],accel_mss,speed_ms,0,blend_radius_m)
  speed_ms = 0.005
  movel([0.204957, -0.671385, -2.812592, -1.228411, 1.570796, 1.775753],accel_mss,speed_ms,0,blend_radius_m)
  speed_ms = 0.040
  movel([0.226788, -0.653095, -2.814511, -1.244783, 1.570796, 1.797585],accel_mss,speed_ms,0,blend_radius_m)
  speed_ms = 0.005
  movel([0.226788, -0.659800, -2.821239, -1.231350, 1.570796, 1.797585],accel_mss,speed_ms,0,blend_radius_m)
  speed_ms = 0.025
  movel([0.226566, -0.650801, -2.822136, -1.239451, 1.570796, 1.797362],accel_mss,speed_ms,0,blend_radius_m)
  movel([0.225962, -0.646853, -2.822519, -1.243016, 1.570796, 1.796758],accel_mss,speed_ms,0,blend_radius_m)
  movel([0.224859, -0.643483, -2.822842, -1.246065, 1.570796, 1.795656],accel_mss,speed_ms,0,blend_radius_m)
  movel([0.223137, -0.640853, -2.823090, -1.248446, 1.570796, 1.793933],accel_mss,speed_ms,0,blend_radius_m)
  movel([0.220667, -0.639133, -2.823251, -1.250005, 1.570796, 1.791464],accel_mss,speed_ms,0,blend_radius_m)
  movel([0.217324, -0.638477, -2.823312, -1.250600, 1.570796, 1.788120],accel_mss,speed_ms,0,blend_radius_m)
  movel([0.212992, -0.639053, -2.823258, -1.250078, 1.570796, 1.783788],accel_mss,speed_ms,0,blend_radius_m)
  speed_ms = 0.005
  movel([0.212992, -0.632672, -2.816490, -1.263228, 1.570796, 1.783788],accel_mss,speed_ms,0,blend_radius_m)
  speed_ms = 0.040
  movel([0.232327, -0.624043, -2.817275, -1.271072, 1.570796, 1.803124],accel_mss,speed_ms,0,blend_radius_m)
  speed_ms = 0.005
  movel([0.232327, -0.630283, -2.824059, -1.258047, 1.570796, 1.803124],accel_mss,speed_ms,0,blend_radius_m)
  speed_ms = 0.025
  movel([0.233592, -0.623885, -2.824625, -1.263880, 1.570796, 1.804388],accel_mss,speed_ms,0,blend_radius_m)
  movel([0.234489, -0.617616, -2.825163, -1.269610, 1.570796, 1.805285],accel_mss,speed_ms,0,blend_radius_m)
  movel([0.234865, -0.611707, -2.825657, -1.275025, 1.570796, 1.805662],accel_mss,speed_ms,0,blend_radius_m)
  movel([0.234575, -0.606409, -2.826087, -1.279893, 1.570796, 1.805371],accel_mss,speed_ms,0,blend_radius_m)
  movel([0.233465, -0.601953, -2.826442, -1.283994, 1.570796, 1.804261],accel_mss,speed_ms,0,blend_radius_m)
  movel([0.232550, -0.600128, -2.826584, -1.285677, 1.570796, 1.803347],accel_mss,speed_ms,0,blend_radius_m)
  movel([0.229927, -0.597415, -2.826794, -1.288179, 1.570796, 1.800723],accel_mss,speed_ms,0,blend_radius_m)
  movel([0.228177, -0.596596, -2.826857, -1.288936, 1.570796, 1.798973],accel_mss,speed_ms,0,blend_radius_m)
  movel([0.226109, -0.596173, -2.826889, -1.289327, 1.570796, 1.796905],accel_mss,speed_ms,0,blend_radius_m)
  movel([0.223710, -0.596181, -2.826889, -1.289319, 1.570796, 1.794507],accel_mss,speed_ms,0,blend_radius_m)
  speed_ms = 0.005
  movel([0.223710, -0.590508, -2.820047, -1.301834, 1.570796, 1.794507],accel_mss,speed_ms,0,blend_radius_m)
  speed_ms = 0.040
  movel([0.244747, -0.579988, -2.820826, -1.311574, 1.570796, 1.815543],accel_mss,speed_ms,0,blend_radius_m)
  speed_ms = 0.005
  movel([0.244747, -0.585477, -2.827685, -1.299227, 1.570796, 1.815543],accel_mss,speed_ms,0,blend_radius_m)
  speed_ms = 0.025
  movel([0.246755, -0.577620, -2.828242, -1.306527, 1.570796, 1.817551],accel_mss,speed_ms,0,blend_radius_m)
  movel([0.248116, -0.570097, -2.828754, -1.313538, 1.570796, 1.818913],accel_mss,speed_ms,0,blend_radius_m)
  movel([0.248691, -0.563170, -2.829206, -1.320013, 1.570796, 1.819487],accel_mss,speed_ms,0,blend_radius_m)
  movel([0.248301, -0.557142, -2.829586, -1.325661, 1.570796, 1.819097],accel_mss,speed_ms,0,blend_radius_m)
  movel([0.246800, -0.552290, -2.829882, -1.330217, 1.570796, 1.817596],accel_mss,speed_ms,0,blend_radius_m)
  movel([0.245573, -0.550405, -2.829995, -1.331990, 1.570796, 1.816369],accel_mss,speed_ms,0,blend_radius_m)
  movel([0.244017, -0.548912, -2.830083, -1.333394, 1.570796, 1.814813],accel_mss,speed_ms,0,blend_radius_m)
  movel([0.242096, -0.547873, -2.830144, -1.334372, 1.570796, 1.812893],accel_mss,speed_ms,0,blend_radius_m)
  movel([0.239802, -0.547300, -2.830178, -1.334911, 1.570796, 1.810599],accel_mss,speed_ms,0,blend_radius_m)
  movel([0.237118, -0.547245, -2.830181, -1.334963, 1.570796, 1.807915],accel_mss,speed_ms,0,blend_radius_m)
  movel([0.234025, -0.547730, -2.830152, -1.334507, 1.570796, 1.804821],accel_mss,speed_ms,0,blend_radius_m)
  speed_ms = 0.005
  movel([0.234025, -0.542915, -2.823242, -1.346232, 1.570796, 1.804821],accel_mss,speed_ms,0,blend_radius_m)
  speed_ms = 0.040
  movel([0.134268, -0.613788, -2.818169, -1.280432, 1.570796, 1.705065],accel_mss,speed_ms,0,blend_radius_m)
  speed_ms = 0.005
  movel([0.134268, -0.619858, -2.824972, -1.267558, 1.570796, 1.705065],accel_mss,speed_ms,0,blend_radius_m)
  speed_ms = 0.025
  movel([0.139062, -0.619665, -2.824989, -1.267735, 1.570796, 1.709858],accel_mss,speed_ms,0,blend_radius_m)
  movel([0.143343, -0.620318, -2.824933, -1.267138, 1.570796, 1.714139],accel_mss,speed_ms,0,blend_radius_m)
  movel([0.147131, -0.621757, -2.824809, -1.265823, 1.570796, 1.717927],accel_mss,speed_ms,0,blend_radius_m)
  movel([0.150438, -0.623920, -2.824622, -1.263847, 1.570796, 1.721234],accel_mss,speed_ms,0,blend_radius_m)
  movel([0.153266, -0.626756, -2.824373, -1.261260, 1.570796, 1.724062],accel_mss,speed_ms,0,blend_radius_m)
  movel([0.155649, -0.630191, -2.824068, -1.258130, 1.570796, 1.726445],accel_mss,speed_ms,0,blend_radius_m)
  movel([0.157585, -0.634180, -2.823707, -1.254502, 1.570796, 1.728381],accel_mss,speed_ms,0,blend_radius_m)
  movel([0.159113, -0.638638, -2.823297, -1.250454, 1.570796, 1.729909],accel_mss,speed_ms,0,blend_radius_m)
  movel([0.160234, -0.643519, -2.822838, -1.246032, 1.570796, 1.731031],accel_mss,speed_ms,0,blend_radius_m)
  movel([0.160985, -0.648749, -2.822336, -1.241303, 1.570796, 1.731782],accel_mss,speed_ms,0,blend_radius_m)
  movel([0.161377, -0.654267, -2.821795, -1.236327, 1.570796, 1.732173],accel_mss,speed_ms,0,blend_radius_m)
  movel([0.161433, -0.660021, -2.821216, -1.231151, 1.570796, 1.732229],accel_mss,speed_ms,0,blend_radius_m)
  movel([0.161176, -0.665932, -2.820608, -1.225848, 1.570796, 1.731972],accel_mss,speed_ms,0,blend_radius_m)
  movel([0.160617, -0.671964, -2.819973, -1.220452, 1.570796, 1.731414],accel_mss,speed_ms,0,blend_radius_m)
  movel([0.159785, -0.678038, -2.819318, -1.215034, 1.570796, 1.730581],accel_mss,speed_ms,0,blend_radius_m)
  movel([0.158700, -0.684106, -2.818648, -1.209635, 1.570796, 1.729497],accel_mss,speed_ms,0,blend_radius_m)
  movel([0.156908, -0.692334, -2.817714, -1.202341, 1.570796, 1.727704],accel_mss,speed_ms,0,blend_radius_m)
  movel([0.154407, -0.701958, -2.816584, -1.193846, 1.570796, 1.725204],accel_mss,speed_ms,0,blend_radius_m)
  movel([0.151119, -0.712273, -2.815329, -1.184787, 1.570796, 1.721915],accel_mss,speed_ms,0,blend_radius_m)
  movel([0.149156, -0.717477, -2.814677, -1.180235, 1.570796, 1.719952],accel_mss,speed_ms,0,blend_radius_m)
  movel([0.146975, -0.722588, -2.814026, -1.175775, 1.570796, 1.717771],accel_mss,speed_ms,0,blend_radius_m)
  movel([0.144549, -0.727547, -2.813383, -1.171459, 1.570796, 1.715345],accel_mss,speed_ms,0,blend_radius_m)
  movel([0.141880, -0.732252, -2.812762, -1.167375, 1.570796, 1.712676],accel_mss,speed_ms,0,blend_radius_m)
  movel([0.138944, -0.736644, -2.812173, -1.163572, 1.570796, 1.709741],accel_mss,speed_ms,0,blend_radius_m)
  movel([0.135729, -0.740650, -2.811628, -1.160111, 1.570796, 1.706525],accel_mss,speed_ms,0,blend_radius_m)
  movel([0.132223, -0.744183, -2.811142, -1.157064, 1.570796, 1.703020],accel_mss,speed_ms,0,blend_radius_m)
  movel([0.128404, -0.747189, -2.810723, -1.154477, 1.570796, 1.699201],accel_mss,speed_ms,0,blend_radius_m)
  movel([0.126366, -0.748472, -2.810543, -1.153374, 1.570796, 1.697163],accel_mss,speed_ms,0,blend_radius_m)
  movel([0.124243, -0.749599, -2.810385, -1.152406, 1.570796, 1.695039],accel_mss,speed_ms,0,blend_radius_m)
  movel([0.119724, -0.751347, -2.810137, -1.150905, 1.570796, 1.690521],accel_mss,speed_ms,0,blend_radius_m)
  movel([0.114551, -0.752607, -2.809958, -1.149824, 1.570796, 1.685347],accel_mss,speed_ms,0,blend_radius_m)
  movel([0.109817, -0.753216, -2.809871, -1.149302, 1.570796, 1.680614],accel_mss,speed_ms,0,blend_radius_m)
  movel([0.105467, -0.753250, -2.809866, -1.149272, 1.570796, 1.676263],accel_mss,speed_ms,0,blend_radius_m)
  movel([0.101426, -0.752776, -2.809934, -1.149679, 1.570796, 1.672223],accel_mss,speed_ms,0,blend_radius_m)
  movel([0.097644, -0.751859, -2.810065, -1.150466, 1.570796, 1.668440],accel_mss,speed_ms,0,blend_radius_m)
  movel([0.094051, -0.750575, -2.810247, -1.151567, 1.570796, 1.664847],accel_mss,speed_ms,0,blend_radius_m)
  movel([0.087186, -0.747177, -2.810725, -1.154487, 1.570796, 1.657982],accel_mss,speed_ms,0,blend_radius_m)
  movel([0.079841, -0.743087, -2.811293, -1.158008, 1.570796, 1.650638],accel_mss,speed_ms,0,blend_radius_m)
  movel([0.072694, -0.738811, -2.811879, -1.161699, 1.570796, 1.643490],accel_mss,speed_ms,0,blend_radius_m)
  movel([0.065973, -0.733946, -2.812536, -1.165907, 1.570796, 1.636769],accel_mss,speed_ms,0,blend_radius_m)
  movel([0.062851, -0.731154, -2.812908, -1.168328, 1.570796, 1.633647],accel_mss,speed_ms,0,blend_radius_m)
  movel([0.059928, -0.728046, -2.813317, -1.171026, 1.570796, 1.630725],accel_mss,speed_ms,0,blend_radius_m)
  movel([0.056167, -0.724321, -2.813802, -1.174265, 1.570796, 1.626963],accel_mss,speed_ms,0,blend_radius_m)
  movel([0.051841, -0.721154, -2.814210, -1.177025, 1.570796, 1.622637],accel_mss,speed_ms,0,blend_radius_m)
  movel([0.047031, -0.718509, -2.814547, -1.179333, 1.570796, 1.617827],accel_mss,speed_ms,0,blend_radius_m)
  movel([0.041837, -0.716319, -2.814823, -1.181246, 1.570796, 1.612633],accel_mss,speed_ms,0,blend_radius_m)
  movel([0.030653, -0.713114, -2.815224, -1.184051, 1.570796, 1.601450],accel_mss,speed_ms,0,blend_radius_m)
  movel([0.019045, -0.711048, -2.815480, -1.185860, 1.570796, 1.589842],accel_mss,speed_ms,0,blend_radius_m)
  movel([0.009832, -0.710334, -2.815568, -1.186487, 1.570796, 1.580628],accel_mss,speed_ms,0,blend_radius_m)
  movel([-0.000049, -0.710772, -2.815514, -1.186103, 1.570796, 1.570748],accel_mss,speed_ms,0,blend_radius_m)
  movel([-0.010548, -0.712385, -2.815315, -1.184689, 1.570796, 1.560248],accel_mss,speed_ms,0,blend_radius_m)
  movel([-0.021606, -0.715202, -2.814964, -1.182224, 1.570796, 1.549190],accel_mss,speed_ms,0,blend_radius_m)
  movel([-0.033162, -0.719217, -2.814457, -1.178715, 1.570796, 1.537634],accel_mss,speed_ms,0,blend_radius_m)
  movel([-0.039102, -0.721676, -2.814143, -1.176570, 1.570796, 1.531694],accel_mss,speed_ms,0,blend_radius_m)
  movel([-0.051271, -0.727491, -2.813390, -1.171508, 1.570796, 1.519526],accel_mss,speed_ms,0,blend_radius_m)
  movel([-0.057482, -0.730846, -2.812948, -1.168594, 1.570796, 1.513315],accel_mss,speed_ms,0,blend_radius_m)
  movel([-0.070094, -0.738431, -2.811931, -1.162027, 1.570796, 1.500702],accel_mss,speed_ms,0,blend_radius_m)
  movel([-0.078788, -0.744355, -2.811118, -1.156916, 1.570796, 1.492008],accel_mss,speed_ms,0,blend_radius_m)
  movel([-0.087499, -0.750990, -2.810188, -1.151211, 1.570796, 1.483298],accel_mss,speed_ms,0,blend_radius_m)
  movel([-0.096132, -0.758258, -2.809145, -1.144985, 1.570796, 1.474664],accel_mss,speed_ms,0,blend_radius_m)
  movel([-0.104601, -0.766099, -2.807992, -1.138298, 1.570796, 1.466195],accel_mss,speed_ms,0,blend_radius_m)
  movel([-0.112827, -0.774447, -2.806731, -1.131210, 1.570796, 1.457969],accel_mss,speed_ms,0,blend_radius_m)
  movel([-0.120726, -0.783232, -2.805368, -1.123789, 1.570796, 1.450070],accel_mss,speed_ms,0,blend_radius_m)
  movel([-0.128222, -0.792392, -2.803905, -1.116092, 1.570796, 1.442574],accel_mss,speed_ms,0,blend_radius_m)
  movel([-0.135243, -0.801861, -2.802348, -1.108180, 1.570796, 1.435553],accel_mss,speed_ms,0,blend_radius_m)
  movel([-0.141321, -0.810835, -2.800831, -1.100724, 1.570796, 1.429476],accel_mss,speed_ms,0,blend_radius_m)
  movel([-0.146733, -0.819572, -2.799312, -1.093505, 1.570796, 1.424064],accel_mss,speed_ms,0,blend_radius_m)
